REGION Network 38: Transition for STATE Num:43 Check Recovery
   RUNG wire#powerrail
      Contact( #s43_ChkRecovery )
      I_Contact( #sStWtResetRel )
      Contact( #sSst )
      wire#w1
      I_Contact( #iProcessOver )
      Coil( #s43_ChkRecovery_T1 )
   END_RUNG
   RUNG wire#w1
      I_Contact( #s43_ChkRecovery_T1 )
      Contact( #iProcessOver )
      Coil( #s43_ChkRecovery_T2 )
   END_RUNG
   // the same network as SCL:
   #_w1 := #s43_ChkRecovery AND NOT #sStWtResetRel AND #sSst;
   #s43_ChkRecovery_T1 := #_w1 AND NOT #iProcessOver;
   #s43_ChkRecovery_T2 := #_w1 AND NOT #s43_ChkRecovery_T1 AND #iProcessOver;
END_REGION

REGION Network 39: STATE Num:43 Check Recovery
   RUNG wire#powerrail
      Contact( #s43_ChkRecovery )
      wire#w1
      I_Contact( #sStWtResetRel )
      I_Contact( #s43_ChkRecovery_T1 )
      I_Contact( #s43_ChkRecovery_T2 )
      wire#w2
      Coil( #s43_ChkRecovery )
   END_RUNG
   RUNG wire#powerrail
      Contact( #s29_WaitProcStart_T1 )
   END_RUNG wire#w1
   RUNG wire#w2
      { S7_GenerateENO := "TRUE" } Move(in := 43, out1 => #StateNo)
   END_RUNG
   // the same network as SCL:
   #s43_ChkRecovery := (#s43_ChkRecovery OR #s29_WaitProcStart_T1) AND NOT #sStWtResetRel AND NOT #s43_ChkRecovery_T1 AND NOT #s43_ChkRecovery_T2;
   IF #s43_ChkRecovery THEN #StateNo := 43; END_IF;
END_REGION
END_FUNCTION_BLOCK

FUNCTION_BLOCK "PR_PC4005_Operator_DecisionV4_653444"   // FB2, LAD
VERSION : 0.1
// stored: AutoNumber true, IsIECCheckEnabled false, UDAEnableTagReadback false
   VAR_INPUT
      iAutoRunning : Bool;
      iOperatorAuthorizationPB : Bool;
      iPCAckZero : Bool;
      iPCBypass : Bool;
      iPCDataReadOver : Bool;
      iPCDataWriteOver : Bool;
      iPalletPresentAtStation : Bool;
      iProcessOver : Bool;
      iProcessStartFormPZR : Bool;
      iRejectPB : Bool;
      iResetMem : Bool;
      iReset_fault : Bool;
      iScanOver : Bool;
      iScanResultNok : Bool;
      iScanResultOk : Bool;
      iScannerBypass : Bool;
      iSstMode : Bool;
      iSstPB : Bool;
      iUnloadCycleSelection : Bool;
   END_VAR
   VAR_OUTPUT
      qPCReadCmd : Bool;
      qPCWriteCmd : Bool;
      qProcessOver : Bool;
      qResetPalletStatusData : Bool;
      qScanCmd : Bool;
   END_VAR
   VAR DB_SPECIFIC
      StateNo : Int;
      s29_WaitProcStart : Bool;
      s29_WaitProcStart_T1 : Bool;
      s30_WaitCartnSheetOp : Bool;
      s30_WaitCartnSheetOp_T1 : Bool;
      s31_ChkCycleSelect : Bool;
      s31_ChkCycleSelect_T1 : Bool;
      s31_ChkCycleSelect_T2 : Bool;
      s32_WaitScanOver : Bool;
      s32_WaitScanOver_T1 : Bool;
      s33_ChkScanResult : Bool;
      s33_ChkScanResult_T1 : Bool;
      s33_ChkScanResult_T2 : Bool;
      s34_WaitOpDecision : Bool;
      s34_WaitOpDecision_T1 : Bool;
      s34_WaitOpDecision_T2 : Bool;
      s35_ChkPCAckReset0 : Bool;
      s35_ChkPCAckReset0_T1 : Bool;
      s36_WaitDataReadPC : Bool;
      s36_WaitDataReadPC_T1 : Bool;
      s38_WaitProcStartLow : Bool;
      s38_WaitProcStartLow_T1 : Bool;
      s39_WaitPalletAbsnt : Bool;
      s39_WaitPalletAbsnt_T1 : Bool;
      s40_WaitFaultReset : Bool;
      s40_WaitFaultReset_T1 : Bool;
      s41_ChkPCAckReset0Up : Bool;
      s41_ChkPCAckReset0Up_T1 : Bool;
      s42_WaitDataUploadPC : Bool;
      s42_WaitDataUploadPC_T1 : Bool;
      s43_ChkRecovery : Bool;
      s43_ChkRecovery_T1 : Bool;
      s43_ChkRecovery_T2 : Bool;
      sPalletAccepted : Bool;
      sProcessOver : Bool;
      sSst : Bool;
      sSstPulse : Bool;
      sSstRise : Bool;
      sStWtResetRel : Bool;
      sStWtResetRel_T1 : Bool;
   END_VAR
   VAR_TEMP
      tOne : Bool;
   END_VAR
   VAR_TEMP   // added for the SCL form of the ladder/FBD networks
      _w1 : Bool;
   END_VAR
BEGIN

REGION Network 1
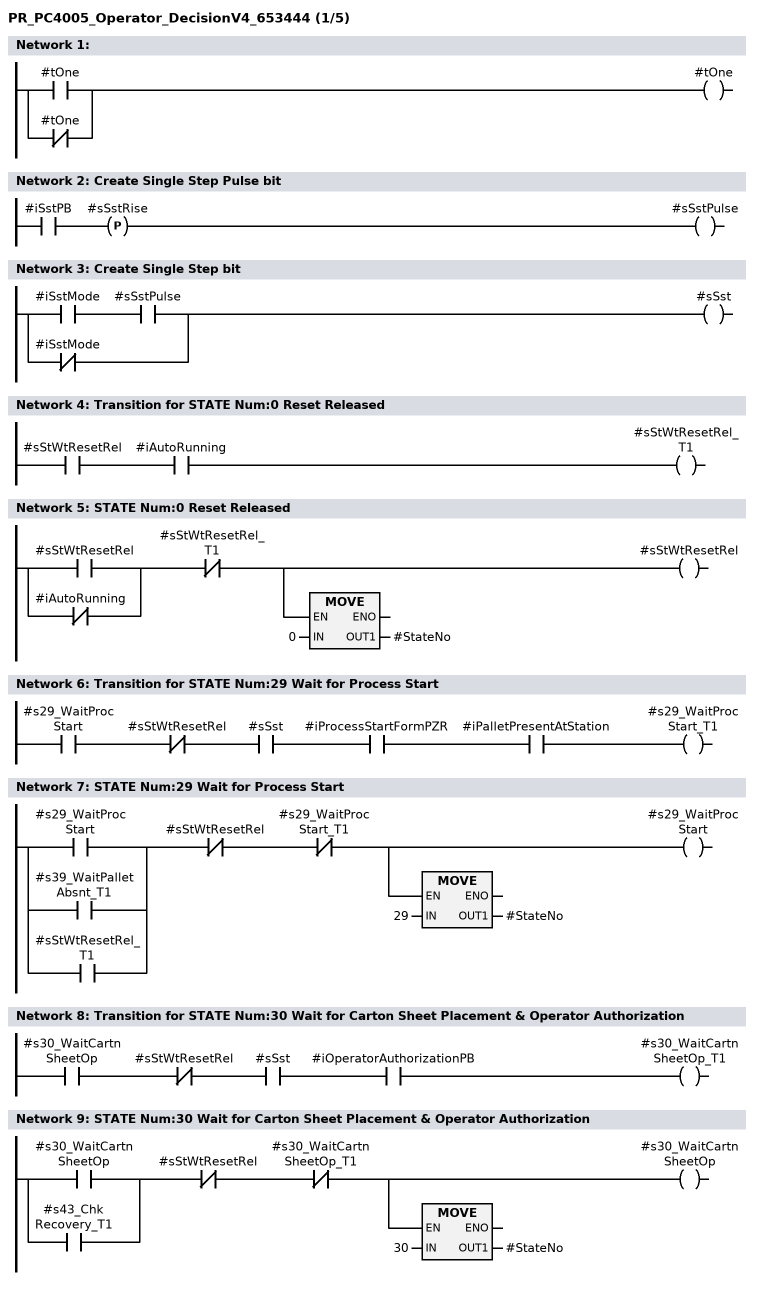
   RUNG wire#powerrail
      Contact( #tOne )
      wire#w1
      Coil( #tOne )
   END_RUNG
   RUNG wire#powerrail
      I_Contact( #tOne )
   END_RUNG wire#w1
   // the same network as SCL:
   #tOne := #tOne OR NOT #tOne;
END_REGION

REGION Network 2: Create Single Step Pulse bit
   RUNG wire#powerrail
      Contact( #iSstPB )
      P_Trig( #sSstRise )
      Coil( #sSstPulse )
   END_RUNG
   // the same network as SCL:
   #_w1 := #iSstPB AND NOT #sSstRise;   // rising edge
   #sSstRise := #iSstPB;
   #sSstPulse := #_w1;
END_REGION

REGION Network 3: Create Single Step bit
   RUNG wire#powerrail
      Contact( #iSstMode )
      Contact( #sSstPulse )
      wire#w1
      Coil( #sSst )
   END_RUNG
   RUNG wire#powerrail
      I_Contact( #iSstMode )
   END_RUNG wire#w1
   // the same network as SCL:
   #sSst := (#iSstMode AND #sSstPulse) OR NOT #iSstMode;
END_REGION

REGION Network 4: Transition for STATE Num:0 Reset Released
   RUNG wire#powerrail
      Contact( #sStWtResetRel )
      Contact( #iAutoRunning )
      Coil( #sStWtResetRel_T1 )
   END_RUNG
   // the same network as SCL:
   #sStWtResetRel_T1 := #sStWtResetRel AND #iAutoRunning;
END_REGION

REGION Network 5: STATE Num:0 Reset Released
   RUNG wire#powerrail
      Contact( #sStWtResetRel )
      wire#w1
      I_Contact( #sStWtResetRel_T1 )
      wire#w2
      Coil( #sStWtResetRel )
   END_RUNG
   RUNG wire#powerrail
      I_Contact( #iAutoRunning )
   END_RUNG wire#w1
   RUNG wire#w2
      { S7_GenerateENO := "TRUE" } Move(in := 0, out1 => #StateNo)
   END_RUNG
   // the same network as SCL:
   #sStWtResetRel := (#sStWtResetRel OR NOT #iAutoRunning) AND NOT #sStWtResetRel_T1;
   IF #sStWtResetRel THEN #StateNo := 0; END_IF;
END_REGION

REGION Network 6: Transition for STATE Num:29 Wait for Process Start
   RUNG wire#powerrail
      Contact( #s29_WaitProcStart )
      I_Contact( #sStWtResetRel )
      Contact( #sSst )
      Contact( #iProcessStartFormPZR )
      Contact( #iPalletPresentAtStation )
      Coil( #s29_WaitProcStart_T1 )
   END_RUNG
   // the same network as SCL:
   #s29_WaitProcStart_T1 := #s29_WaitProcStart AND NOT #sStWtResetRel AND #sSst AND #iProcessStartFormPZR AND #iPalletPresentAtStation;
END_REGION

REGION Network 7: STATE Num:29 Wait for Process Start
   RUNG wire#powerrail
      Contact( #s29_WaitProcStart )
      wire#w1
      I_Contact( #sStWtResetRel )
      I_Contact( #s29_WaitProcStart_T1 )
      wire#w2
      Coil( #s29_WaitProcStart )
   END_RUNG
   RUNG wire#powerrail
      Contact( #s39_WaitPalletAbsnt_T1 )
   END_RUNG wire#w1
   RUNG wire#powerrail
      Contact( #sStWtResetRel_T1 )
   END_RUNG wire#w1
   RUNG wire#w2
      { S7_GenerateENO := "TRUE" } Move(in := 29, out1 => #StateNo)
   END_RUNG
   // the same network as SCL:
   #s29_WaitProcStart := (#s29_WaitProcStart OR #s39_WaitPalletAbsnt_T1 OR #sStWtResetRel_T1) AND NOT #sStWtResetRel AND NOT #s29_WaitProcStart_T1;
   IF #s29_WaitProcStart THEN #StateNo := 29; END_IF;
END_REGION

REGION Network 8: Transition for STATE Num:30 Wait for Carton Sheet Placement & Operator Authorization
   RUNG wire#powerrail
      Contact( #s30_WaitCartnSheetOp )
      I_Contact( #sStWtResetRel )
      Contact( #sSst )
      Contact( #iOperatorAuthorizationPB )
      Coil( #s30_WaitCartnSheetOp_T1 )
   END_RUNG
   // the same network as SCL:
   #s30_WaitCartnSheetOp_T1 := #s30_WaitCartnSheetOp AND NOT #sStWtResetRel AND #sSst AND #iOperatorAuthorizationPB;
END_REGION

REGION Network 9: STATE Num:30 Wait for Carton Sheet Placement & Operator Authorization
   RUNG wire#powerrail
      Contact( #s30_WaitCartnSheetOp )
      wire#w1
      I_Contact( #sStWtResetRel )
      I_Contact( #s30_WaitCartnSheetOp_T1 )
      wire#w2
      Coil( #s30_WaitCartnSheetOp )
   END_RUNG
   RUNG wire#powerrail
      Contact( #s43_ChkRecovery_T1 )
   END_RUNG wire#w1
   RUNG wire#w2
      { S7_GenerateENO := "TRUE" } Move(in := 30, out1 => #StateNo)
   END_RUNG
   // the same network as SCL:
   #s30_WaitCartnSheetOp := (#s30_WaitCartnSheetOp OR #s43_ChkRecovery_T1) AND NOT #sStWtResetRel AND NOT #s30_WaitCartnSheetOp_T1;
   IF #s30_WaitCartnSheetOp THEN #StateNo := 30; END_IF;
END_REGION

REGION Network 10: Transition for STATE Num:31 Check Cycle Selection
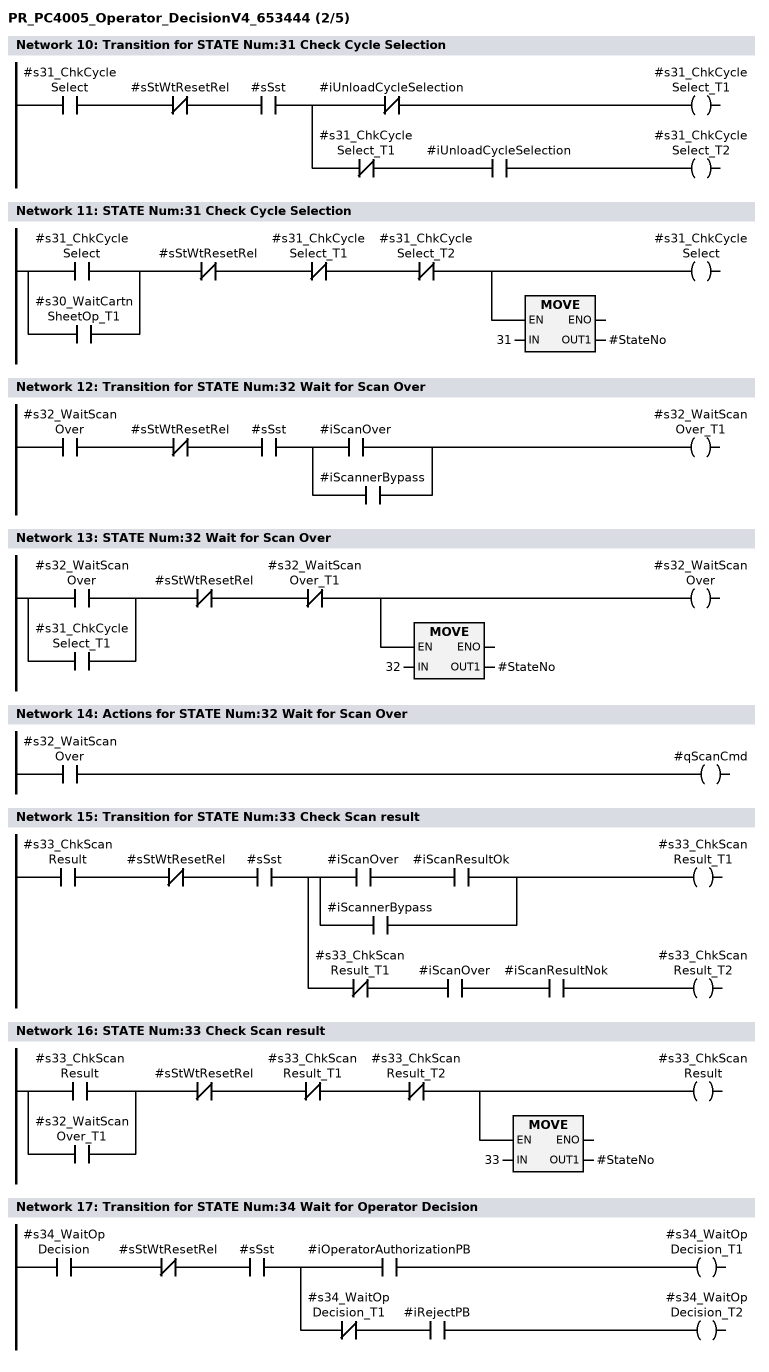
   RUNG wire#powerrail
      Contact( #s31_ChkCycleSelect )
      I_Contact( #sStWtResetRel )
      Contact( #sSst )
      wire#w1
      I_Contact( #iUnloadCycleSelection )
      Coil( #s31_ChkCycleSelect_T1 )
   END_RUNG
   RUNG wire#w1
      I_Contact( #s31_ChkCycleSelect_T1 )
      Contact( #iUnloadCycleSelection )
      Coil( #s31_ChkCycleSelect_T2 )
   END_RUNG
   // the same network as SCL:
   #_w1 := #s31_ChkCycleSelect AND NOT #sStWtResetRel AND #sSst;
   #s31_ChkCycleSelect_T1 := #_w1 AND NOT #iUnloadCycleSelection;
   #s31_ChkCycleSelect_T2 := #_w1 AND NOT #s31_ChkCycleSelect_T1 AND #iUnloadCycleSelection;
END_REGION

REGION Network 11: STATE Num:31 Check Cycle Selection
   RUNG wire#powerrail
      Contact( #s31_ChkCycleSelect )
      wire#w1
      I_Contact( #sStWtResetRel )
      I_Contact( #s31_ChkCycleSelect_T1 )
      I_Contact( #s31_ChkCycleSelect_T2 )
      wire#w2
      Coil( #s31_ChkCycleSelect )
   END_RUNG
   RUNG wire#powerrail
      Contact( #s30_WaitCartnSheetOp_T1 )
   END_RUNG wire#w1
   RUNG wire#w2
      { S7_GenerateENO := "TRUE" } Move(in := 31, out1 => #StateNo)
   END_RUNG
   // the same network as SCL:
   #s31_ChkCycleSelect := (#s31_ChkCycleSelect OR #s30_WaitCartnSheetOp_T1) AND NOT #sStWtResetRel AND NOT #s31_ChkCycleSelect_T1 AND NOT #s31_ChkCycleSelect_T2;
   IF #s31_ChkCycleSelect THEN #StateNo := 31; END_IF;
END_REGION

REGION Network 12: Transition for STATE Num:32 Wait for Scan Over
   RUNG wire#powerrail
      Contact( #s32_WaitScanOver )
      I_Contact( #sStWtResetRel )
      Contact( #sSst )
      wire#w1
      Contact( #iScanOver )
      wire#w2
      Coil( #s32_WaitScanOver_T1 )
   END_RUNG
   RUNG wire#w1
      Contact( #iScannerBypass )
   END_RUNG wire#w2
   // the same network as SCL:
   #s32_WaitScanOver_T1 := #s32_WaitScanOver AND NOT #sStWtResetRel AND #sSst AND (#iScanOver OR #iScannerBypass);
END_REGION

REGION Network 13: STATE Num:32 Wait for Scan Over
   RUNG wire#powerrail
      Contact( #s32_WaitScanOver )
      wire#w1
      I_Contact( #sStWtResetRel )
      I_Contact( #s32_WaitScanOver_T1 )
      wire#w2
      Coil( #s32_WaitScanOver )
   END_RUNG
   RUNG wire#powerrail
      Contact( #s31_ChkCycleSelect_T1 )
   END_RUNG wire#w1
   RUNG wire#w2
      { S7_GenerateENO := "TRUE" } Move(in := 32, out1 => #StateNo)
   END_RUNG
   // the same network as SCL:
   #s32_WaitScanOver := (#s32_WaitScanOver OR #s31_ChkCycleSelect_T1) AND NOT #sStWtResetRel AND NOT #s32_WaitScanOver_T1;
   IF #s32_WaitScanOver THEN #StateNo := 32; END_IF;
END_REGION

REGION Network 14: Actions for STATE Num:32 Wait for Scan Over
   RUNG wire#powerrail
      Contact( #s32_WaitScanOver )
      Coil( #qScanCmd )
   END_RUNG
   // the same network as SCL:
   #qScanCmd := #s32_WaitScanOver;
END_REGION

REGION Network 15: Transition for STATE Num:33 Check Scan result
   RUNG wire#powerrail
      Contact( #s33_ChkScanResult )
      I_Contact( #sStWtResetRel )
      Contact( #sSst )
      wire#w1
      Contact( #iScanOver )
      Contact( #iScanResultOk )
      wire#w2
      Coil( #s33_ChkScanResult_T1 )
   END_RUNG
   RUNG wire#w1
      Contact( #iScannerBypass )
   END_RUNG wire#w2
   RUNG wire#w1
      I_Contact( #s33_ChkScanResult_T1 )
      Contact( #iScanOver )
      Contact( #iScanResultNok )
      Coil( #s33_ChkScanResult_T2 )
   END_RUNG
   // the same network as SCL:
   #_w1 := #s33_ChkScanResult AND NOT #sStWtResetRel AND #sSst;
   #s33_ChkScanResult_T1 := #_w1 AND ((#iScanOver AND #iScanResultOk) OR #iScannerBypass);
   #s33_ChkScanResult_T2 := #_w1 AND NOT #s33_ChkScanResult_T1 AND #iScanOver AND #iScanResultNok;
END_REGION

REGION Network 16: STATE Num:33 Check Scan result
   RUNG wire#powerrail
      Contact( #s33_ChkScanResult )
      wire#w1
      I_Contact( #sStWtResetRel )
      I_Contact( #s33_ChkScanResult_T1 )
      I_Contact( #s33_ChkScanResult_T2 )
      wire#w2
      Coil( #s33_ChkScanResult )
   END_RUNG
   RUNG wire#powerrail
      Contact( #s32_WaitScanOver_T1 )
   END_RUNG wire#w1
   RUNG wire#w2
      { S7_GenerateENO := "TRUE" } Move(in := 33, out1 => #StateNo)
   END_RUNG
   // the same network as SCL:
   #s33_ChkScanResult := (#s33_ChkScanResult OR #s32_WaitScanOver_T1) AND NOT #sStWtResetRel AND NOT #s33_ChkScanResult_T1 AND NOT #s33_ChkScanResult_T2;
   IF #s33_ChkScanResult THEN #StateNo := 33; END_IF;
END_REGION

REGION Network 17: Transition for STATE Num:34 Wait for Operator Decision
   RUNG wire#powerrail
      Contact( #s34_WaitOpDecision )
      I_Contact( #sStWtResetRel )
      Contact( #sSst )
      wire#w1
      Contact( #iOperatorAuthorizationPB )
      Coil( #s34_WaitOpDecision_T1 )
   END_RUNG
   RUNG wire#w1
      I_Contact( #s34_WaitOpDecision_T1 )
      Contact( #iRejectPB )
      Coil( #s34_WaitOpDecision_T2 )
   END_RUNG
   // the same network as SCL:
   #_w1 := #s34_WaitOpDecision AND NOT #sStWtResetRel AND #sSst;
   #s34_WaitOpDecision_T1 := #_w1 AND #iOperatorAuthorizationPB;
   #s34_WaitOpDecision_T2 := #_w1 AND NOT #s34_WaitOpDecision_T1 AND #iRejectPB;
END_REGION

REGION Network 18: STATE Num:34 Wait for Operator Decision
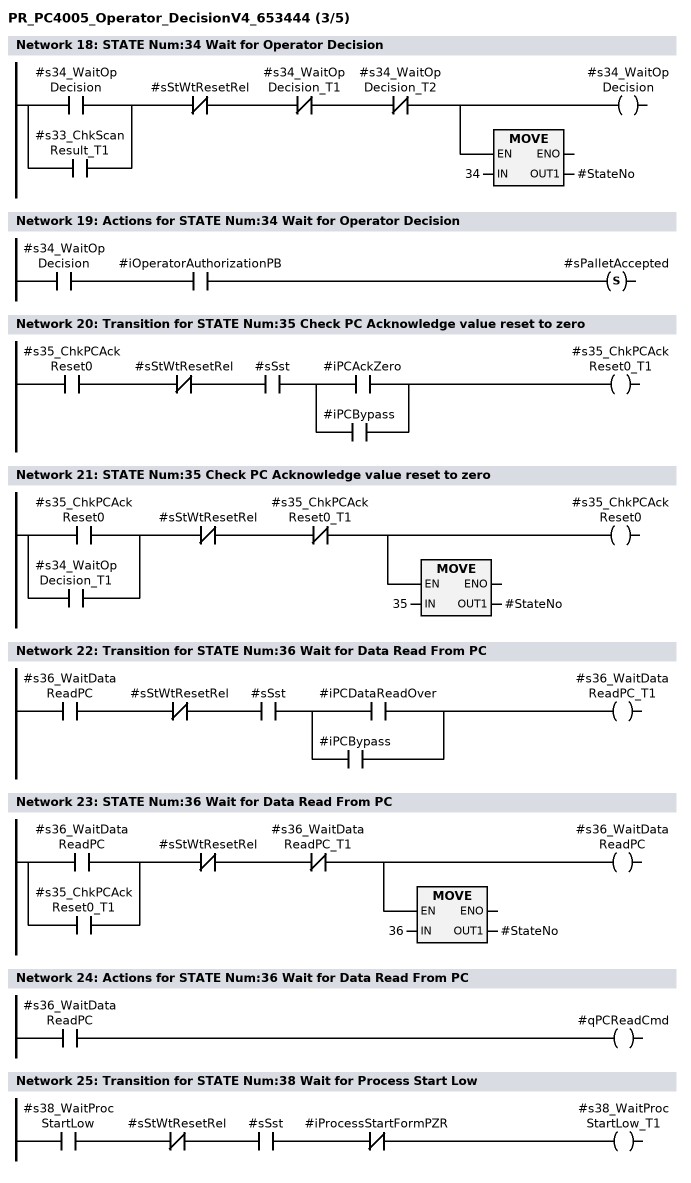
   RUNG wire#powerrail
      Contact( #s34_WaitOpDecision )
      wire#w1
      I_Contact( #sStWtResetRel )
      I_Contact( #s34_WaitOpDecision_T1 )
      I_Contact( #s34_WaitOpDecision_T2 )
      wire#w2
      Coil( #s34_WaitOpDecision )
   END_RUNG
   RUNG wire#powerrail
      Contact( #s33_ChkScanResult_T1 )
   END_RUNG wire#w1
   RUNG wire#w2
      { S7_GenerateENO := "TRUE" } Move(in := 34, out1 => #StateNo)
   END_RUNG
   // the same network as SCL:
   #s34_WaitOpDecision := (#s34_WaitOpDecision OR #s33_ChkScanResult_T1) AND NOT #sStWtResetRel AND NOT #s34_WaitOpDecision_T1 AND NOT #s34_WaitOpDecision_T2;
   IF #s34_WaitOpDecision THEN #StateNo := 34; END_IF;
END_REGION

REGION Network 19: Actions for STATE Num:34 Wait for Operator Decision
   RUNG wire#powerrail
      Contact( #s34_WaitOpDecision )
      Contact( #iOperatorAuthorizationPB )
      S_Coil( #sPalletAccepted )
   END_RUNG
   // the same network as SCL:
   IF #s34_WaitOpDecision AND #iOperatorAuthorizationPB THEN #sPalletAccepted := TRUE; END_IF;
END_REGION

REGION Network 20: Transition for STATE Num:35 Check PC Acknowledge value reset to zero
   RUNG wire#powerrail
      Contact( #s35_ChkPCAckReset0 )
      I_Contact( #sStWtResetRel )
      Contact( #sSst )
      wire#w1
      Contact( #iPCAckZero )
      wire#w2
      Coil( #s35_ChkPCAckReset0_T1 )
   END_RUNG
   RUNG wire#w1
      Contact( #iPCBypass )
   END_RUNG wire#w2
   // the same network as SCL:
   #s35_ChkPCAckReset0_T1 := #s35_ChkPCAckReset0 AND NOT #sStWtResetRel AND #sSst AND (#iPCAckZero OR #iPCBypass);
END_REGION

REGION Network 21: STATE Num:35 Check PC Acknowledge value reset to zero
   RUNG wire#powerrail
      Contact( #s35_ChkPCAckReset0 )
      wire#w1
      I_Contact( #sStWtResetRel )
      I_Contact( #s35_ChkPCAckReset0_T1 )
      wire#w2
      Coil( #s35_ChkPCAckReset0 )
   END_RUNG
   RUNG wire#powerrail
      Contact( #s34_WaitOpDecision_T1 )
   END_RUNG wire#w1
   RUNG wire#w2
      { S7_GenerateENO := "TRUE" } Move(in := 35, out1 => #StateNo)
   END_RUNG
   // the same network as SCL:
   #s35_ChkPCAckReset0 := (#s35_ChkPCAckReset0 OR #s34_WaitOpDecision_T1) AND NOT #sStWtResetRel AND NOT #s35_ChkPCAckReset0_T1;
   IF #s35_ChkPCAckReset0 THEN #StateNo := 35; END_IF;
END_REGION

REGION Network 22: Transition for STATE Num:36 Wait for Data Read From PC
   RUNG wire#powerrail
      Contact( #s36_WaitDataReadPC )
      I_Contact( #sStWtResetRel )
      Contact( #sSst )
      wire#w1
      Contact( #iPCDataReadOver )
      wire#w2
      Coil( #s36_WaitDataReadPC_T1 )
   END_RUNG
   RUNG wire#w1
      Contact( #iPCBypass )
   END_RUNG wire#w2
   // the same network as SCL:
   #s36_WaitDataReadPC_T1 := #s36_WaitDataReadPC AND NOT #sStWtResetRel AND #sSst AND (#iPCDataReadOver OR #iPCBypass);
END_REGION

REGION Network 23: STATE Num:36 Wait for Data Read From PC
   RUNG wire#powerrail
      Contact( #s36_WaitDataReadPC )
      wire#w1
      I_Contact( #sStWtResetRel )
      I_Contact( #s36_WaitDataReadPC_T1 )
      wire#w2
      Coil( #s36_WaitDataReadPC )
   END_RUNG
   RUNG wire#powerrail
      Contact( #s35_ChkPCAckReset0_T1 )
   END_RUNG wire#w1
   RUNG wire#w2
      { S7_GenerateENO := "TRUE" } Move(in := 36, out1 => #StateNo)
   END_RUNG
   // the same network as SCL:
   #s36_WaitDataReadPC := (#s36_WaitDataReadPC OR #s35_ChkPCAckReset0_T1) AND NOT #sStWtResetRel AND NOT #s36_WaitDataReadPC_T1;
   IF #s36_WaitDataReadPC THEN #StateNo := 36; END_IF;
END_REGION

REGION Network 24: Actions for STATE Num:36 Wait for Data Read From PC
   RUNG wire#powerrail
      Contact( #s36_WaitDataReadPC )
      Coil( #qPCReadCmd )
   END_RUNG
   // the same network as SCL:
   #qPCReadCmd := #s36_WaitDataReadPC;
END_REGION

REGION Network 25: Transition for STATE Num:38 Wait for Process Start Low
   RUNG wire#powerrail
      Contact( #s38_WaitProcStartLow )
      I_Contact( #sStWtResetRel )
      Contact( #sSst )
      I_Contact( #iProcessStartFormPZR )
      Coil( #s38_WaitProcStartLow_T1 )
   END_RUNG
   // the same network as SCL:
   #s38_WaitProcStartLow_T1 := #s38_WaitProcStartLow AND NOT #sStWtResetRel AND #sSst AND NOT #iProcessStartFormPZR;
END_REGION

REGION Network 26: STATE Num:38 Wait for Process Start Low
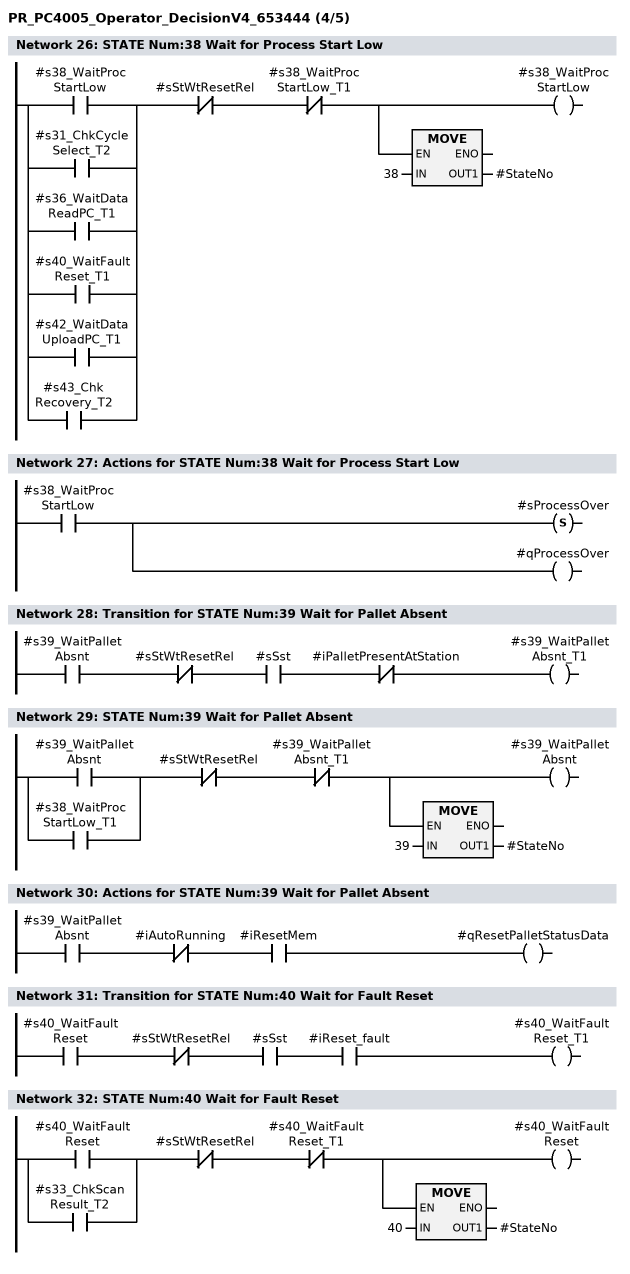
   RUNG wire#powerrail
      Contact( #s38_WaitProcStartLow )
      wire#w1
      I_Contact( #sStWtResetRel )
      I_Contact( #s38_WaitProcStartLow_T1 )
      wire#w2
      Coil( #s38_WaitProcStartLow )
   END_RUNG
   RUNG wire#powerrail
      Contact( #s31_ChkCycleSelect_T2 )
   END_RUNG wire#w1
   RUNG wire#powerrail
      Contact( #s36_WaitDataReadPC_T1 )
   END_RUNG wire#w1
   RUNG wire#powerrail
      Contact( #s40_WaitFaultReset_T1 )
   END_RUNG wire#w1
   RUNG wire#powerrail
      Contact( #s42_WaitDataUploadPC_T1 )
   END_RUNG wire#w1
   RUNG wire#powerrail
      Contact( #s43_ChkRecovery_T2 )
   END_RUNG wire#w1
   RUNG wire#w2
      { S7_GenerateENO := "TRUE" } Move(in := 38, out1 => #StateNo)
   END_RUNG
   // the same network as SCL:
   #s38_WaitProcStartLow := (#s38_WaitProcStartLow OR #s31_ChkCycleSelect_T2 OR #s36_WaitDataReadPC_T1 OR #s40_WaitFaultReset_T1 OR #s42_WaitDataUploadPC_T1 OR #s43_ChkRecovery_T2) AND NOT #sStWtResetRel AND NOT #s38_WaitProcStartLow_T1;
   IF #s38_WaitProcStartLow THEN #StateNo := 38; END_IF;
END_REGION

REGION Network 27: Actions for STATE Num:38 Wait for Process Start Low
   RUNG wire#powerrail
      Contact( #s38_WaitProcStartLow )
      wire#w1
      S_Coil( #sProcessOver )
   END_RUNG
   RUNG wire#w1
      Coil( #qProcessOver )
   END_RUNG
   // the same network as SCL:
   IF #s38_WaitProcStartLow THEN #sProcessOver := TRUE; END_IF;
   #qProcessOver := #s38_WaitProcStartLow;
END_REGION

REGION Network 28: Transition for STATE Num:39 Wait for Pallet Absent
   RUNG wire#powerrail
      Contact( #s39_WaitPalletAbsnt )
      I_Contact( #sStWtResetRel )
      Contact( #sSst )
      I_Contact( #iPalletPresentAtStation )
      Coil( #s39_WaitPalletAbsnt_T1 )
   END_RUNG
   // the same network as SCL:
   #s39_WaitPalletAbsnt_T1 := #s39_WaitPalletAbsnt AND NOT #sStWtResetRel AND #sSst AND NOT #iPalletPresentAtStation;
END_REGION

REGION Network 29: STATE Num:39 Wait for Pallet Absent
   RUNG wire#powerrail
      Contact( #s39_WaitPalletAbsnt )
      wire#w1
      I_Contact( #sStWtResetRel )
      I_Contact( #s39_WaitPalletAbsnt_T1 )
      wire#w2
      Coil( #s39_WaitPalletAbsnt )
   END_RUNG
   RUNG wire#powerrail
      Contact( #s38_WaitProcStartLow_T1 )
   END_RUNG wire#w1
   RUNG wire#w2
      { S7_GenerateENO := "TRUE" } Move(in := 39, out1 => #StateNo)
   END_RUNG
   // the same network as SCL:
   #s39_WaitPalletAbsnt := (#s39_WaitPalletAbsnt OR #s38_WaitProcStartLow_T1) AND NOT #sStWtResetRel AND NOT #s39_WaitPalletAbsnt_T1;
   IF #s39_WaitPalletAbsnt THEN #StateNo := 39; END_IF;
END_REGION

REGION Network 30: Actions for STATE Num:39 Wait for Pallet Absent
   RUNG wire#powerrail
      Contact( #s39_WaitPalletAbsnt )
      I_Contact( #iAutoRunning )
      Contact( #iResetMem )
      Coil( #qResetPalletStatusData )
   END_RUNG
   // the same network as SCL:
   #qResetPalletStatusData := #s39_WaitPalletAbsnt AND NOT #iAutoRunning AND #iResetMem;
END_REGION

REGION Network 31: Transition for STATE Num:40 Wait for Fault Reset
   RUNG wire#powerrail
      Contact( #s40_WaitFaultReset )
      I_Contact( #sStWtResetRel )
      Contact( #sSst )
      Contact( #iReset_fault )
      Coil( #s40_WaitFaultReset_T1 )
   END_RUNG
   // the same network as SCL:
   #s40_WaitFaultReset_T1 := #s40_WaitFaultReset AND NOT #sStWtResetRel AND #sSst AND #iReset_fault;
END_REGION

REGION Network 32: STATE Num:40 Wait for Fault Reset
   RUNG wire#powerrail
      Contact( #s40_WaitFaultReset )
      wire#w1
      I_Contact( #sStWtResetRel )
      I_Contact( #s40_WaitFaultReset_T1 )
      wire#w2
      Coil( #s40_WaitFaultReset )
   END_RUNG
   RUNG wire#powerrail
      Contact( #s33_ChkScanResult_T2 )
   END_RUNG wire#w1
   RUNG wire#w2
      { S7_GenerateENO := "TRUE" } Move(in := 40, out1 => #StateNo)
   END_RUNG
   // the same network as SCL:
   #s40_WaitFaultReset := (#s40_WaitFaultReset OR #s33_ChkScanResult_T2) AND NOT #sStWtResetRel AND NOT #s40_WaitFaultReset_T1;
   IF #s40_WaitFaultReset THEN #StateNo := 40; END_IF;
END_REGION

REGION Network 33: Transition for STATE Num:41 Check PC Acknowledge value reset to zero for Upload
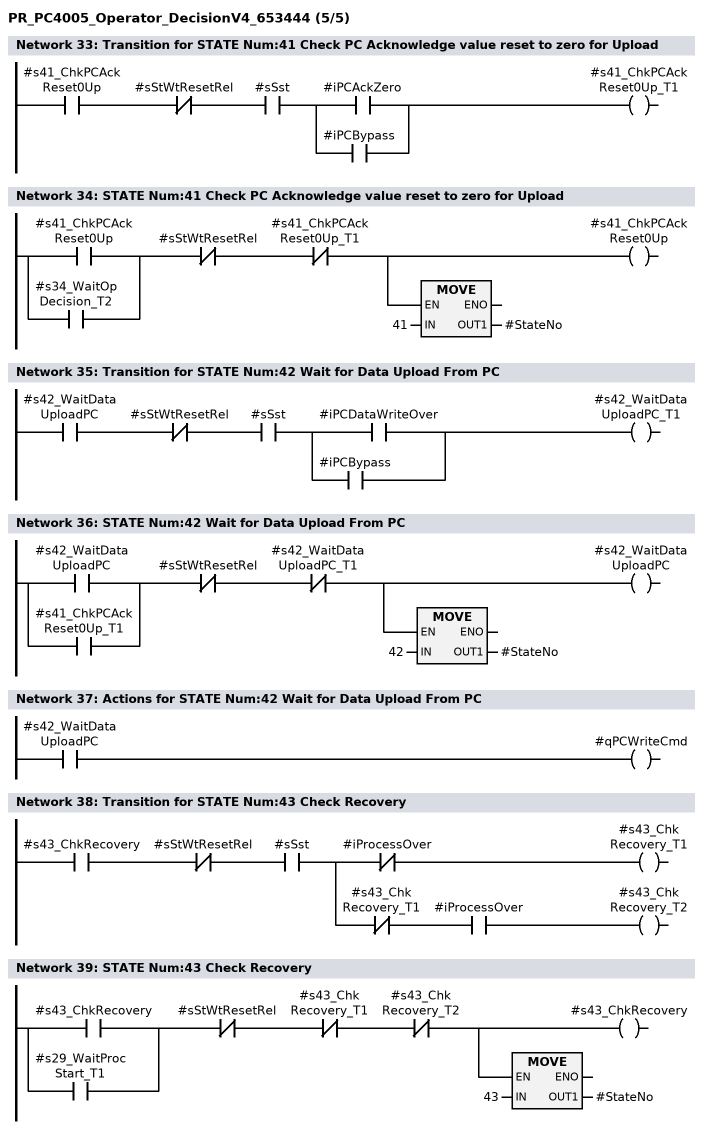
   RUNG wire#powerrail
      Contact( #s41_ChkPCAckReset0Up )
      I_Contact( #sStWtResetRel )
      Contact( #sSst )
      wire#w1
      Contact( #iPCAckZero )
      wire#w2
      Coil( #s41_ChkPCAckReset0Up_T1 )
   END_RUNG
   RUNG wire#w1
      Contact( #iPCBypass )
   END_RUNG wire#w2
   // the same network as SCL:
   #s41_ChkPCAckReset0Up_T1 := #s41_ChkPCAckReset0Up AND NOT #sStWtResetRel AND #sSst AND (#iPCAckZero OR #iPCBypass);
END_REGION

REGION Network 34: STATE Num:41 Check PC Acknowledge value reset to zero for Upload
   RUNG wire#powerrail
      Contact( #s41_ChkPCAckReset0Up )
      wire#w1
      I_Contact( #sStWtResetRel )
      I_Contact( #s41_ChkPCAckReset0Up_T1 )
      wire#w2
      Coil( #s41_ChkPCAckReset0Up )
   END_RUNG
   RUNG wire#powerrail
      Contact( #s34_WaitOpDecision_T2 )
   END_RUNG wire#w1
   RUNG wire#w2
      { S7_GenerateENO := "TRUE" } Move(in := 41, out1 => #StateNo)
   END_RUNG
   // the same network as SCL:
   #s41_ChkPCAckReset0Up := (#s41_ChkPCAckReset0Up OR #s34_WaitOpDecision_T2) AND NOT #sStWtResetRel AND NOT #s41_ChkPCAckReset0Up_T1;
   IF #s41_ChkPCAckReset0Up THEN #StateNo := 41; END_IF;
END_REGION

REGION Network 35: Transition for STATE Num:42 Wait for Data Upload From PC
   RUNG wire#powerrail
      Contact( #s42_WaitDataUploadPC )
      I_Contact( #sStWtResetRel )
      Contact( #sSst )
      wire#w1
      Contact( #iPCDataWriteOver )
      wire#w2
      Coil( #s42_WaitDataUploadPC_T1 )
   END_RUNG
   RUNG wire#w1
      Contact( #iPCBypass )
   END_RUNG wire#w2
   // the same network as SCL:
   #s42_WaitDataUploadPC_T1 := #s42_WaitDataUploadPC AND NOT #sStWtResetRel AND #sSst AND (#iPCDataWriteOver OR #iPCBypass);
END_REGION

REGION Network 36: STATE Num:42 Wait for Data Upload From PC
   RUNG wire#powerrail
      Contact( #s42_WaitDataUploadPC )
      wire#w1
      I_Contact( #sStWtResetRel )
      I_Contact( #s42_WaitDataUploadPC_T1 )
      wire#w2
      Coil( #s42_WaitDataUploadPC )
   END_RUNG
   RUNG wire#powerrail
      Contact( #s41_ChkPCAckReset0Up_T1 )
   END_RUNG wire#w1
   RUNG wire#w2
      { S7_GenerateENO := "TRUE" } Move(in := 42, out1 => #StateNo)
   END_RUNG
   // the same network as SCL:
   #s42_WaitDataUploadPC := (#s42_WaitDataUploadPC OR #s41_ChkPCAckReset0Up_T1) AND NOT #sStWtResetRel AND NOT #s42_WaitDataUploadPC_T1;
   IF #s42_WaitDataUploadPC THEN #StateNo := 42; END_IF;
END_REGION

REGION Network 37: Actions for STATE Num:42 Wait for Data Upload From PC
   RUNG wire#powerrail
      Contact( #s42_WaitDataUploadPC )
      Coil( #qPCWriteCmd )
   END_RUNG
   // the same network as SCL:
   #qPCWriteCmd := #s42_WaitDataUploadPC;
END_REGION

REGION Network 38: Transition for STATE Num:43 Check Recovery
   RUNG wire#powerrail
      Contact( #s43_ChkRecovery )
      I_Contact( #sStWtResetRel )
      Contact( #sSst )
      wire#w1
      I_Contact( #iProcessOver )
      Coil( #s43_ChkRecovery_T1 )
   END_RUNG
   RUNG wire#w1
      I_Contact( #s43_ChkRecovery_T1 )
      Contact( #iProcessOver )
      Coil( #s43_ChkRecovery_T2 )
   END_RUNG
   // the same network as SCL:
   #_w1 := #s43_ChkRecovery AND NOT #sStWtResetRel AND #sSst;
   #s43_ChkRecovery_T1 := #_w1 AND NOT #iProcessOver;
   #s43_ChkRecovery_T2 := #_w1 AND NOT #s43_ChkRecovery_T1 AND #iProcessOver;
END_REGION

REGION Network 39: STATE Num:43 Check Recovery
   RUNG wire#powerrail
      Contact( #s43_ChkRecovery )
      wire#w1
      I_Contact( #sStWtResetRel )
      I_Contact( #s43_ChkRecovery_T1 )
      I_Contact( #s43_ChkRecovery_T2 )
      wire#w2
      Coil( #s43_ChkRecovery )
   END_RUNG
   RUNG wire#powerrail
      Contact( #s29_WaitProcStart_T1 )
   END_RUNG wire#w1
   RUNG wire#w2
      { S7_GenerateENO := "TRUE" } Move(in := 43, out1 => #StateNo)
   END_RUNG
   // the same network as SCL:
   #s43_ChkRecovery := (#s43_ChkRecovery OR #s29_WaitProcStart_T1) AND NOT #sStWtResetRel AND NOT #s43_ChkRecovery_T1 AND NOT #s43_ChkRecovery_T2;
   IF #s43_ChkRecovery THEN #StateNo := 43; END_IF;
END_REGION
END_FUNCTION_BLOCK

FUNCTION_BLOCK "PR_PC4005_Operator_DecisionV4_77a371"   // FB1, LAD
VERSION : 0.1
// stored: AutoNumber true, IsIECCheckEnabled false, UDAEnableTagReadback false
   VAR_INPUT
      iAutoRunning : Bool;
      iOperatorAuthorizationPB : Bool;
      iPCAckZero : Bool;
      iPCBypass : Bool;
      iPCDataReadOver : Bool;
      iPCDataWriteOver : Bool;
      iPalletPresentAtStation : Bool;
      iProcessOver : Bool;
      iProcessStartFormPZR : Bool;
      iRejectPB : Bool;
      iResetMem : Bool;
      iReset_fault : Bool;
      iScanOver : Bool;
      iScanResultNok : Bool;
      iScanResultOk : Bool;
      iScannerBypass : Bool;
      iSstMode : Bool;
      iSstPB : Bool;
      iUnloadCycleSelection : Bool;
   END_VAR
   VAR_OUTPUT
      qPCReadCmd : Bool;
      qPCWriteCmd : Bool;
      qProcessOver : Bool;
      qResetPalletStatusData : Bool;
      qScanCmd : Bool;
   END_VAR
   VAR DB_SPECIFIC
      StateNo : Int;
      s29_WaitProcStart : Bool;
      s29_WaitProcStart_T1 : Bool;
      s30_WaitCartnSheetOp : Bool;
      s30_WaitCartnSheetOp_T1 : Bool;
      s31_ChkCycleSelect : Bool;
      s31_ChkCycleSelect_T1 : Bool;
      s31_ChkCycleSelect_T2 : Bool;
      s32_WaitScanOver : Bool;
      s32_WaitScanOver_T1 : Bool;
      s33_ChkScanResult : Bool;
      s33_ChkScanResult_T1 : Bool;
      s33_ChkScanResult_T2 : Bool;
      s34_WaitOpDecision : Bool;
      s34_WaitOpDecision_T1 : Bool;
      s34_WaitOpDecision_T2 : Bool;
      s35_ChkPCAckReset0 : Bool;
      s35_ChkPCAckReset0_T1 : Bool;
      s36_WaitDataReadPC : Bool;
      s36_WaitDataReadPC_T1 : Bool;
      s38_WaitProcStartLow : Bool;
      s38_WaitProcStartLow_T1 : Bool;
      s39_WaitPalletAbsnt : Bool;
      s39_WaitPalletAbsnt_T1 : Bool;
      s40_WaitFaultReset : Bool;
      s40_WaitFaultReset_T1 : Bool;
      s41_ChkPCAckReset0Up : Bool;
      s41_ChkPCAckReset0Up_T1 : Bool;
      s42_WaitDataUploadPC : Bool;
      s42_WaitDataUploadPC_T1 : Bool;
      s43_ChkRecovery : Bool;
      s43_ChkRecovery_T1 : Bool;
      s43_ChkRecovery_T2 : Bool;
      sPalletAccepted : Bool;
      sProcessOver : Bool;
      sSst : Bool;
      sSstPulse : Bool;
      sSstRise : Bool;
      sStWtResetRel : Bool;
      sStWtResetRel_T1 : Bool;
   END_VAR
   VAR_TEMP
      tOne : Bool;
   END_VAR
   VAR_TEMP   // added for the SCL form of the ladder/FBD networks
      _w1 : Bool;
   END_VAR
BEGIN

REGION Network 1
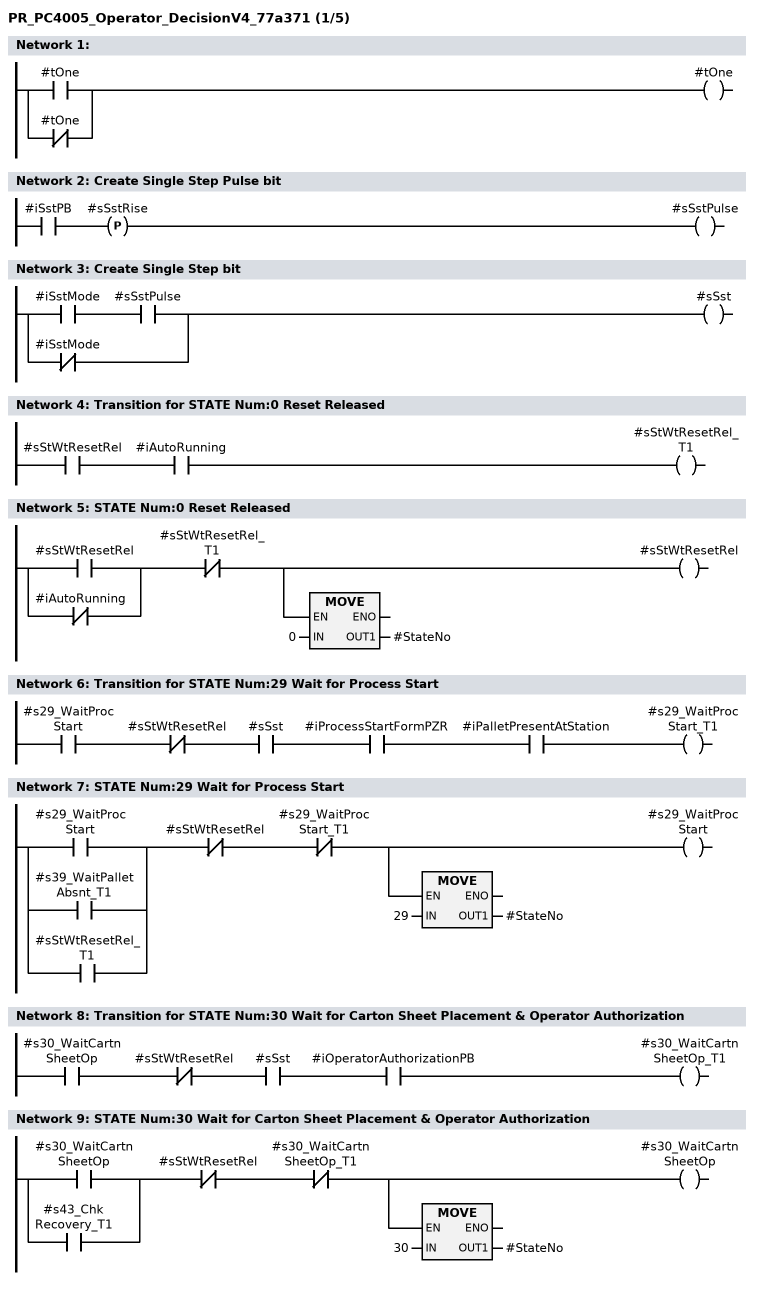
   RUNG wire#powerrail
      Contact( #tOne )
      wire#w1
      Coil( #tOne )
   END_RUNG
   RUNG wire#powerrail
      I_Contact( #tOne )
   END_RUNG wire#w1
   // the same network as SCL:
   #tOne := #tOne OR NOT #tOne;
END_REGION

REGION Network 2: Create Single Step Pulse bit
   RUNG wire#powerrail
      Contact( #iSstPB )
      P_Trig( #sSstRise )
      Coil( #sSstPulse )
   END_RUNG
   // the same network as SCL:
   #_w1 := #iSstPB AND NOT #sSstRise;   // rising edge
   #sSstRise := #iSstPB;
   #sSstPulse := #_w1;
END_REGION

REGION Network 3: Create Single Step bit
   RUNG wire#powerrail
      Contact( #iSstMode )
      Contact( #sSstPulse )
      wire#w1
      Coil( #sSst )
   END_RUNG
   RUNG wire#powerrail
      I_Contact( #iSstMode )
   END_RUNG wire#w1
   // the same network as SCL:
   #sSst := (#iSstMode AND #sSstPulse) OR NOT #iSstMode;
END_REGION

REGION Network 4: Transition for STATE Num:0 Reset Released
   RUNG wire#powerrail
      Contact( #sStWtResetRel )
      Contact( #iAutoRunning )
      Coil( #sStWtResetRel_T1 )
   END_RUNG
   // the same network as SCL:
   #sStWtResetRel_T1 := #sStWtResetRel AND #iAutoRunning;
END_REGION

REGION Network 5: STATE Num:0 Reset Released
   RUNG wire#powerrail
      Contact( #sStWtResetRel )
      wire#w1
      I_Contact( #sStWtResetRel_T1 )
      wire#w2
      Coil( #sStWtResetRel )
   END_RUNG
   RUNG wire#powerrail
      I_Contact( #iAutoRunning )
   END_RUNG wire#w1
   RUNG wire#w2
      { S7_GenerateENO := "TRUE" } Move(in := 0, out1 => #StateNo)
   END_RUNG
   // the same network as SCL:
   #sStWtResetRel := (#sStWtResetRel OR NOT #iAutoRunning) AND NOT #sStWtResetRel_T1;
   IF #sStWtResetRel THEN #StateNo := 0; END_IF;
END_REGION

REGION Network 6: Transition for STATE Num:29 Wait for Process Start
   RUNG wire#powerrail
      Contact( #s29_WaitProcStart )
      I_Contact( #sStWtResetRel )
      Contact( #sSst )
      Contact( #iProcessStartFormPZR )
      Contact( #iPalletPresentAtStation )
      Coil( #s29_WaitProcStart_T1 )
   END_RUNG
   // the same network as SCL:
   #s29_WaitProcStart_T1 := #s29_WaitProcStart AND NOT #sStWtResetRel AND #sSst AND #iProcessStartFormPZR AND #iPalletPresentAtStation;
END_REGION

REGION Network 7: STATE Num:29 Wait for Process Start
   RUNG wire#powerrail
      Contact( #s29_WaitProcStart )
      wire#w1
      I_Contact( #sStWtResetRel )
      I_Contact( #s29_WaitProcStart_T1 )
      wire#w2
      Coil( #s29_WaitProcStart )
   END_RUNG
   RUNG wire#powerrail
      Contact( #s39_WaitPalletAbsnt_T1 )
   END_RUNG wire#w1
   RUNG wire#powerrail
      Contact( #sStWtResetRel_T1 )
   END_RUNG wire#w1
   RUNG wire#w2
      { S7_GenerateENO := "TRUE" } Move(in := 29, out1 => #StateNo)
   END_RUNG
   // the same network as SCL:
   #s29_WaitProcStart := (#s29_WaitProcStart OR #s39_WaitPalletAbsnt_T1 OR #sStWtResetRel_T1) AND NOT #sStWtResetRel AND NOT #s29_WaitProcStart_T1;
   IF #s29_WaitProcStart THEN #StateNo := 29; END_IF;
END_REGION

REGION Network 8: Transition for STATE Num:30 Wait for Carton Sheet Placement & Operator Authorization
   RUNG wire#powerrail
      Contact( #s30_WaitCartnSheetOp )
      I_Contact( #sStWtResetRel )
      Contact( #sSst )
      Contact( #iOperatorAuthorizationPB )
      Coil( #s30_WaitCartnSheetOp_T1 )
   END_RUNG
   // the same network as SCL:
   #s30_WaitCartnSheetOp_T1 := #s30_WaitCartnSheetOp AND NOT #sStWtResetRel AND #sSst AND #iOperatorAuthorizationPB;
END_REGION

REGION Network 9: STATE Num:30 Wait for Carton Sheet Placement & Operator Authorization
   RUNG wire#powerrail
      Contact( #s30_WaitCartnSheetOp )
      wire#w1
      I_Contact( #sStWtResetRel )
      I_Contact( #s30_WaitCartnSheetOp_T1 )
      wire#w2
      Coil( #s30_WaitCartnSheetOp )
   END_RUNG
   RUNG wire#powerrail
      Contact( #s43_ChkRecovery_T1 )
   END_RUNG wire#w1
   RUNG wire#w2
      { S7_GenerateENO := "TRUE" } Move(in := 30, out1 => #StateNo)
   END_RUNG
   // the same network as SCL:
   #s30_WaitCartnSheetOp := (#s30_WaitCartnSheetOp OR #s43_ChkRecovery_T1) AND NOT #sStWtResetRel AND NOT #s30_WaitCartnSheetOp_T1;
   IF #s30_WaitCartnSheetOp THEN #StateNo := 30; END_IF;
END_REGION

REGION Network 10: Transition for STATE Num:31 Check Cycle Selection
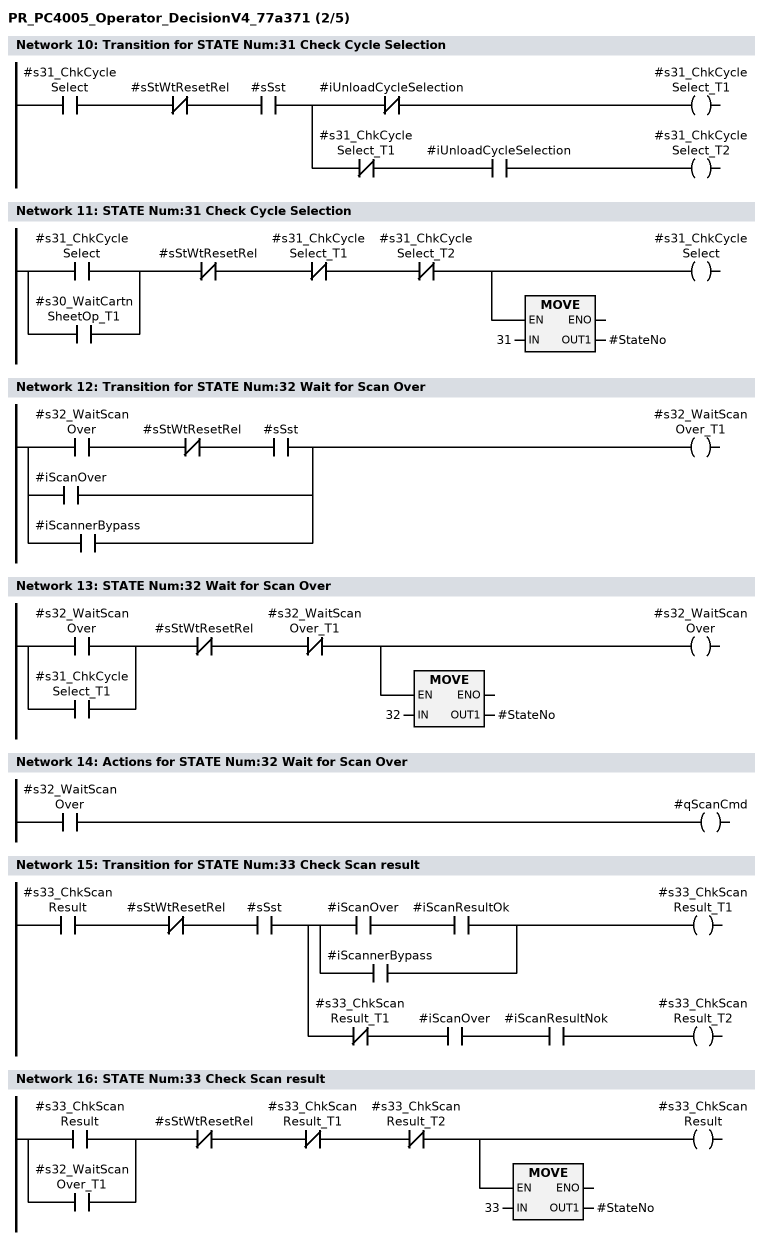
   RUNG wire#powerrail
      Contact( #s31_ChkCycleSelect )
      I_Contact( #sStWtResetRel )
      Contact( #sSst )
      wire#w1
      I_Contact( #iUnloadCycleSelection )
      Coil( #s31_ChkCycleSelect_T1 )
   END_RUNG
   RUNG wire#w1
      I_Contact( #s31_ChkCycleSelect_T1 )
      Contact( #iUnloadCycleSelection )
      Coil( #s31_ChkCycleSelect_T2 )
   END_RUNG
   // the same network as SCL:
   #_w1 := #s31_ChkCycleSelect AND NOT #sStWtResetRel AND #sSst;
   #s31_ChkCycleSelect_T1 := #_w1 AND NOT #iUnloadCycleSelection;
   #s31_ChkCycleSelect_T2 := #_w1 AND NOT #s31_ChkCycleSelect_T1 AND #iUnloadCycleSelection;
END_REGION

REGION Network 11: STATE Num:31 Check Cycle Selection
   RUNG wire#powerrail
      Contact( #s31_ChkCycleSelect )
      wire#w1
      I_Contact( #sStWtResetRel )
      I_Contact( #s31_ChkCycleSelect_T1 )
      I_Contact( #s31_ChkCycleSelect_T2 )
      wire#w2
      Coil( #s31_ChkCycleSelect )
   END_RUNG
   RUNG wire#powerrail
      Contact( #s30_WaitCartnSheetOp_T1 )
   END_RUNG wire#w1
   RUNG wire#w2
      { S7_GenerateENO := "TRUE" } Move(in := 31, out1 => #StateNo)
   END_RUNG
   // the same network as SCL:
   #s31_ChkCycleSelect := (#s31_ChkCycleSelect OR #s30_WaitCartnSheetOp_T1) AND NOT #sStWtResetRel AND NOT #s31_ChkCycleSelect_T1 AND NOT #s31_ChkCycleSelect_T2;
   IF #s31_ChkCycleSelect THEN #StateNo := 31; END_IF;
END_REGION

REGION Network 12: Transition for STATE Num:32 Wait for Scan Over
   RUNG wire#powerrail
      Contact( #s32_WaitScanOver )
      I_Contact( #sStWtResetRel )
      Contact( #sSst )
      wire#w1
      Coil( #s32_WaitScanOver_T1 )
   END_RUNG
   RUNG wire#powerrail
      Contact( #iScanOver )
   END_RUNG wire#w1
   RUNG wire#powerrail
      Contact( #iScannerBypass )
   END_RUNG wire#w1
   // the same network as SCL:
   #s32_WaitScanOver_T1 := (#s32_WaitScanOver AND NOT #sStWtResetRel AND #sSst) OR #iScanOver OR #iScannerBypass;
END_REGION

REGION Network 13: STATE Num:32 Wait for Scan Over
   RUNG wire#powerrail
      Contact( #s32_WaitScanOver )
      wire#w1
      I_Contact( #sStWtResetRel )
      I_Contact( #s32_WaitScanOver_T1 )
      wire#w2
      Coil( #s32_WaitScanOver )
   END_RUNG
   RUNG wire#powerrail
      Contact( #s31_ChkCycleSelect_T1 )
   END_RUNG wire#w1
   RUNG wire#w2
      { S7_GenerateENO := "TRUE" } Move(in := 32, out1 => #StateNo)
   END_RUNG
   // the same network as SCL:
   #s32_WaitScanOver := (#s32_WaitScanOver OR #s31_ChkCycleSelect_T1) AND NOT #sStWtResetRel AND NOT #s32_WaitScanOver_T1;
   IF #s32_WaitScanOver THEN #StateNo := 32; END_IF;
END_REGION

REGION Network 14: Actions for STATE Num:32 Wait for Scan Over
   RUNG wire#powerrail
      Contact( #s32_WaitScanOver )
      Coil( #qScanCmd )
   END_RUNG
   // the same network as SCL:
   #qScanCmd := #s32_WaitScanOver;
END_REGION

REGION Network 15: Transition for STATE Num:33 Check Scan result
   RUNG wire#powerrail
      Contact( #s33_ChkScanResult )
      I_Contact( #sStWtResetRel )
      Contact( #sSst )
      wire#w1
      Contact( #iScanOver )
      Contact( #iScanResultOk )
      wire#w2
      Coil( #s33_ChkScanResult_T1 )
   END_RUNG
   RUNG wire#w1
      Contact( #iScannerBypass )
   END_RUNG wire#w2
   RUNG wire#w1
      I_Contact( #s33_ChkScanResult_T1 )
      Contact( #iScanOver )
      Contact( #iScanResultNok )
      Coil( #s33_ChkScanResult_T2 )
   END_RUNG
   // the same network as SCL:
   #_w1 := #s33_ChkScanResult AND NOT #sStWtResetRel AND #sSst;
   #s33_ChkScanResult_T1 := #_w1 AND ((#iScanOver AND #iScanResultOk) OR #iScannerBypass);
   #s33_ChkScanResult_T2 := #_w1 AND NOT #s33_ChkScanResult_T1 AND #iScanOver AND #iScanResultNok;
END_REGION

REGION Network 16: STATE Num:33 Check Scan result
   RUNG wire#powerrail
      Contact( #s33_ChkScanResult )
      wire#w1
      I_Contact( #sStWtResetRel )
      I_Contact( #s33_ChkScanResult_T1 )
      I_Contact( #s33_ChkScanResult_T2 )
      wire#w2
      Coil( #s33_ChkScanResult )
   END_RUNG
   RUNG wire#powerrail
      Contact( #s32_WaitScanOver_T1 )
   END_RUNG wire#w1
   RUNG wire#w2
      { S7_GenerateENO := "TRUE" } Move(in := 33, out1 => #StateNo)
   END_RUNG
   // the same network as SCL:
   #s33_ChkScanResult := (#s33_ChkScanResult OR #s32_WaitScanOver_T1) AND NOT #sStWtResetRel AND NOT #s33_ChkScanResult_T1 AND NOT #s33_ChkScanResult_T2;
   IF #s33_ChkScanResult THEN #StateNo := 33; END_IF;
END_REGION

REGION Network 17: Transition for STATE Num:34 Wait for Operator Decision
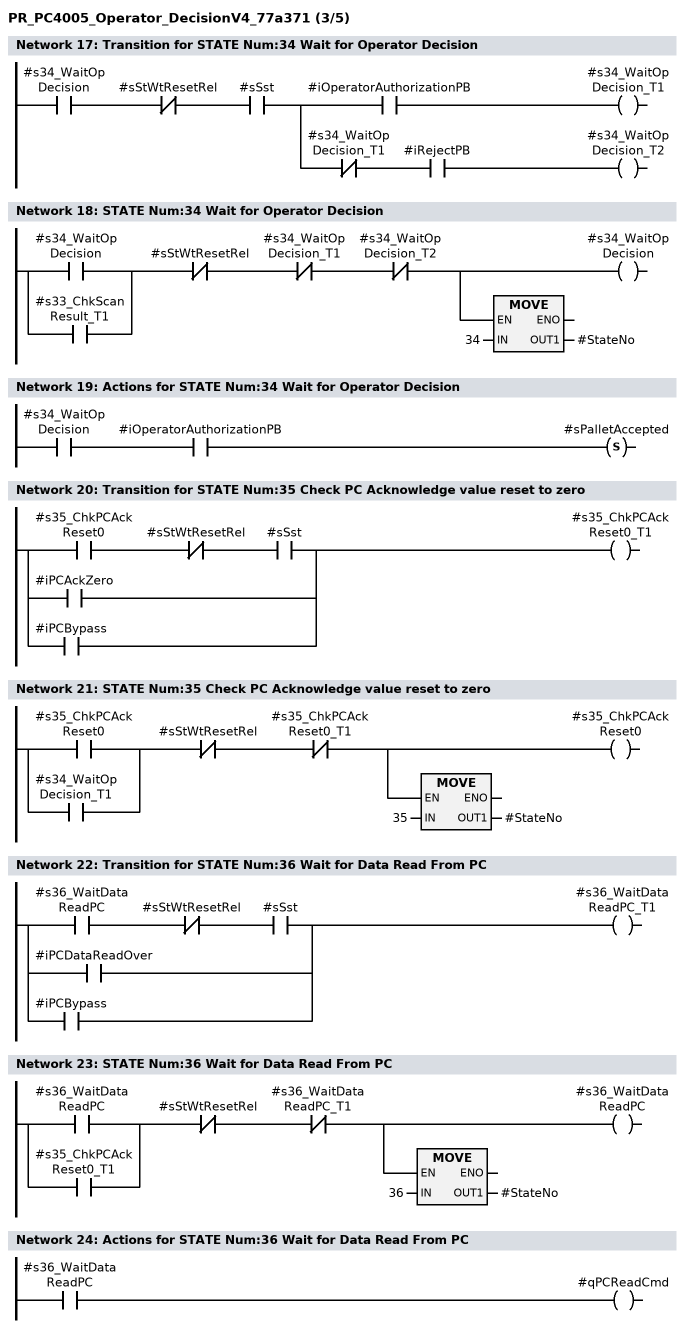
   RUNG wire#powerrail
      Contact( #s34_WaitOpDecision )
      I_Contact( #sStWtResetRel )
      Contact( #sSst )
      wire#w1
      Contact( #iOperatorAuthorizationPB )
      Coil( #s34_WaitOpDecision_T1 )
   END_RUNG
   RUNG wire#w1
      I_Contact( #s34_WaitOpDecision_T1 )
      Contact( #iRejectPB )
      Coil( #s34_WaitOpDecision_T2 )
   END_RUNG
   // the same network as SCL:
   #_w1 := #s34_WaitOpDecision AND NOT #sStWtResetRel AND #sSst;
   #s34_WaitOpDecision_T1 := #_w1 AND #iOperatorAuthorizationPB;
   #s34_WaitOpDecision_T2 := #_w1 AND NOT #s34_WaitOpDecision_T1 AND #iRejectPB;
END_REGION

REGION Network 18: STATE Num:34 Wait for Operator Decision
   RUNG wire#powerrail
      Contact( #s34_WaitOpDecision )
      wire#w1
      I_Contact( #sStWtResetRel )
      I_Contact( #s34_WaitOpDecision_T1 )
      I_Contact( #s34_WaitOpDecision_T2 )
      wire#w2
      Coil( #s34_WaitOpDecision )
   END_RUNG
   RUNG wire#powerrail
      Contact( #s33_ChkScanResult_T1 )
   END_RUNG wire#w1
   RUNG wire#w2
      { S7_GenerateENO := "TRUE" } Move(in := 34, out1 => #StateNo)
   END_RUNG
   // the same network as SCL:
   #s34_WaitOpDecision := (#s34_WaitOpDecision OR #s33_ChkScanResult_T1) AND NOT #sStWtResetRel AND NOT #s34_WaitOpDecision_T1 AND NOT #s34_WaitOpDecision_T2;
   IF #s34_WaitOpDecision THEN #StateNo := 34; END_IF;
END_REGION

REGION Network 19: Actions for STATE Num:34 Wait for Operator Decision
   RUNG wire#powerrail
      Contact( #s34_WaitOpDecision )
      Contact( #iOperatorAuthorizationPB )
      S_Coil( #sPalletAccepted )
   END_RUNG
   // the same network as SCL:
   IF #s34_WaitOpDecision AND #iOperatorAuthorizationPB THEN #sPalletAccepted := TRUE; END_IF;
END_REGION

REGION Network 20: Transition for STATE Num:35 Check PC Acknowledge value reset to zero
   RUNG wire#powerrail
      Contact( #s35_ChkPCAckReset0 )
      I_Contact( #sStWtResetRel )
      Contact( #sSst )
      wire#w1
      Coil( #s35_ChkPCAckReset0_T1 )
   END_RUNG
   RUNG wire#powerrail
      Contact( #iPCAckZero )
   END_RUNG wire#w1
   RUNG wire#powerrail
      Contact( #iPCBypass )
   END_RUNG wire#w1
   // the same network as SCL:
   #s35_ChkPCAckReset0_T1 := (#s35_ChkPCAckReset0 AND NOT #sStWtResetRel AND #sSst) OR #iPCAckZero OR #iPCBypass;
END_REGION

REGION Network 21: STATE Num:35 Check PC Acknowledge value reset to zero
   RUNG wire#powerrail
      Contact( #s35_ChkPCAckReset0 )
      wire#w1
      I_Contact( #sStWtResetRel )
      I_Contact( #s35_ChkPCAckReset0_T1 )
      wire#w2
      Coil( #s35_ChkPCAckReset0 )
   END_RUNG
   RUNG wire#powerrail
      Contact( #s34_WaitOpDecision_T1 )
   END_RUNG wire#w1
   RUNG wire#w2
      { S7_GenerateENO := "TRUE" } Move(in := 35, out1 => #StateNo)
   END_RUNG
   // the same network as SCL:
   #s35_ChkPCAckReset0 := (#s35_ChkPCAckReset0 OR #s34_WaitOpDecision_T1) AND NOT #sStWtResetRel AND NOT #s35_ChkPCAckReset0_T1;
   IF #s35_ChkPCAckReset0 THEN #StateNo := 35; END_IF;
END_REGION

REGION Network 22: Transition for STATE Num:36 Wait for Data Read From PC
   RUNG wire#powerrail
      Contact( #s36_WaitDataReadPC )
      I_Contact( #sStWtResetRel )
      Contact( #sSst )
      wire#w1
      Coil( #s36_WaitDataReadPC_T1 )
   END_RUNG
   RUNG wire#powerrail
      Contact( #iPCDataReadOver )
   END_RUNG wire#w1
   RUNG wire#powerrail
      Contact( #iPCBypass )
   END_RUNG wire#w1
   // the same network as SCL:
   #s36_WaitDataReadPC_T1 := (#s36_WaitDataReadPC AND NOT #sStWtResetRel AND #sSst) OR #iPCDataReadOver OR #iPCBypass;
END_REGION

REGION Network 23: STATE Num:36 Wait for Data Read From PC
   RUNG wire#powerrail
      Contact( #s36_WaitDataReadPC )
      wire#w1
      I_Contact( #sStWtResetRel )
      I_Contact( #s36_WaitDataReadPC_T1 )
      wire#w2
      Coil( #s36_WaitDataReadPC )
   END_RUNG
   RUNG wire#powerrail
      Contact( #s35_ChkPCAckReset0_T1 )
   END_RUNG wire#w1
   RUNG wire#w2
      { S7_GenerateENO := "TRUE" } Move(in := 36, out1 => #StateNo)
   END_RUNG
   // the same network as SCL:
   #s36_WaitDataReadPC := (#s36_WaitDataReadPC OR #s35_ChkPCAckReset0_T1) AND NOT #sStWtResetRel AND NOT #s36_WaitDataReadPC_T1;
   IF #s36_WaitDataReadPC THEN #StateNo := 36; END_IF;
END_REGION

REGION Network 24: Actions for STATE Num:36 Wait for Data Read From PC
   RUNG wire#powerrail
      Contact( #s36_WaitDataReadPC )
      Coil( #qPCReadCmd )
   END_RUNG
   // the same network as SCL:
   #qPCReadCmd := #s36_WaitDataReadPC;
END_REGION

REGION Network 25: Transition for STATE Num:38 Wait for Process Start Low
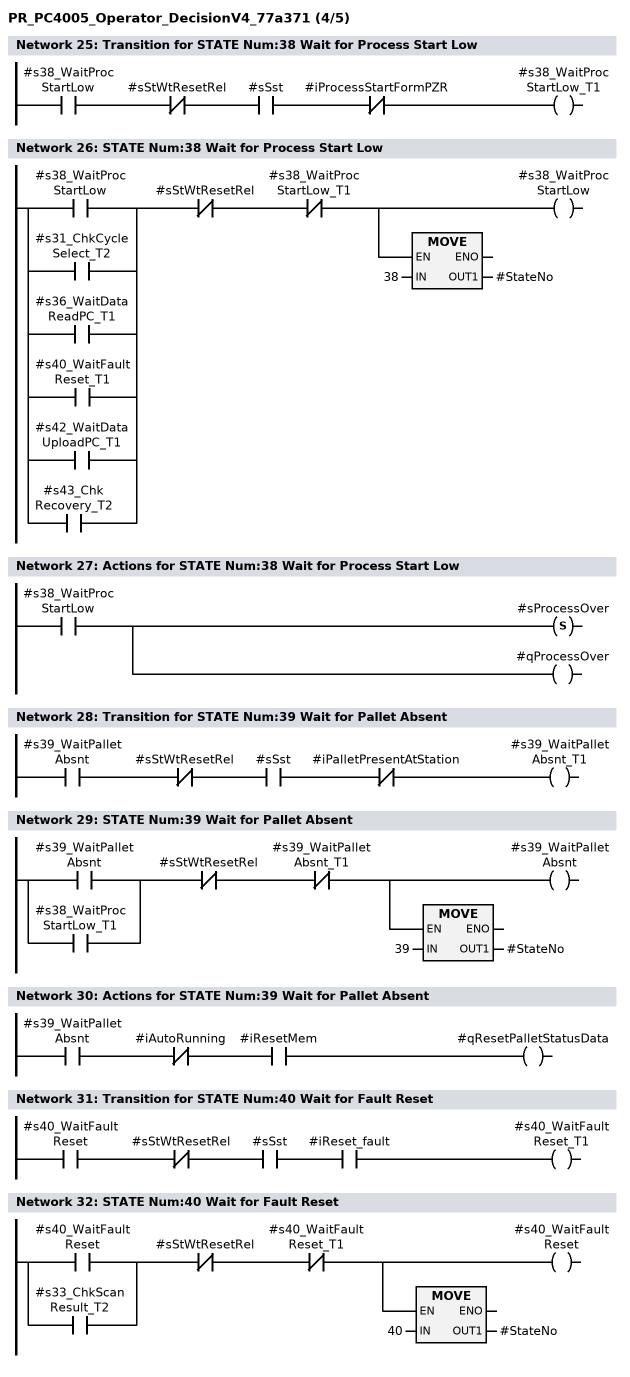
   RUNG wire#powerrail
      Contact( #s38_WaitProcStartLow )
      I_Contact( #sStWtResetRel )
      Contact( #sSst )
      I_Contact( #iProcessStartFormPZR )
      Coil( #s38_WaitProcStartLow_T1 )
   END_RUNG
   // the same network as SCL:
   #s38_WaitProcStartLow_T1 := #s38_WaitProcStartLow AND NOT #sStWtResetRel AND #sSst AND NOT #iProcessStartFormPZR;
END_REGION

REGION Network 26: STATE Num:38 Wait for Process Start Low
   RUNG wire#powerrail
      Contact( #s38_WaitProcStartLow )
      wire#w1
      I_Contact( #sStWtResetRel )
      I_Contact( #s38_WaitProcStartLow_T1 )
      wire#w2
      Coil( #s38_WaitProcStartLow )
   END_RUNG
   RUNG wire#powerrail
      Contact( #s31_ChkCycleSelect_T2 )
   END_RUNG wire#w1
   RUNG wire#powerrail
      Contact( #s36_WaitDataReadPC_T1 )
   END_RUNG wire#w1
   RUNG wire#powerrail
      Contact( #s40_WaitFaultReset_T1 )
   END_RUNG wire#w1
   RUNG wire#powerrail
      Contact( #s42_WaitDataUploadPC_T1 )
   END_RUNG wire#w1
   RUNG wire#powerrail
      Contact( #s43_ChkRecovery_T2 )
   END_RUNG wire#w1
   RUNG wire#w2
      { S7_GenerateENO := "TRUE" } Move(in := 38, out1 => #StateNo)
   END_RUNG
   // the same network as SCL:
   #s38_WaitProcStartLow := (#s38_WaitProcStartLow OR #s31_ChkCycleSelect_T2 OR #s36_WaitDataReadPC_T1 OR #s40_WaitFaultReset_T1 OR #s42_WaitDataUploadPC_T1 OR #s43_ChkRecovery_T2) AND NOT #sStWtResetRel AND NOT #s38_WaitProcStartLow_T1;
   IF #s38_WaitProcStartLow THEN #StateNo := 38; END_IF;
END_REGION

REGION Network 27: Actions for STATE Num:38 Wait for Process Start Low
   RUNG wire#powerrail
      Contact( #s38_WaitProcStartLow )
      wire#w1
      S_Coil( #sProcessOver )
   END_RUNG
   RUNG wire#w1
      Coil( #qProcessOver )
   END_RUNG
   // the same network as SCL:
   IF #s38_WaitProcStartLow THEN #sProcessOver := TRUE; END_IF;
   #qProcessOver := #s38_WaitProcStartLow;
END_REGION

REGION Network 28: Transition for STATE Num:39 Wait for Pallet Absent
   RUNG wire#powerrail
      Contact( #s39_WaitPalletAbsnt )
      I_Contact( #sStWtResetRel )
      Contact( #sSst )
      I_Contact( #iPalletPresentAtStation )
      Coil( #s39_WaitPalletAbsnt_T1 )
   END_RUNG
   // the same network as SCL:
   #s39_WaitPalletAbsnt_T1 := #s39_WaitPalletAbsnt AND NOT #sStWtResetRel AND #sSst AND NOT #iPalletPresentAtStation;
END_REGION

REGION Network 29: STATE Num:39 Wait for Pallet Absent
   RUNG wire#powerrail
      Contact( #s39_WaitPalletAbsnt )
      wire#w1
      I_Contact( #sStWtResetRel )
      I_Contact( #s39_WaitPalletAbsnt_T1 )
      wire#w2
      Coil( #s39_WaitPalletAbsnt )
   END_RUNG
   RUNG wire#powerrail
      Contact( #s38_WaitProcStartLow_T1 )
   END_RUNG wire#w1
   RUNG wire#w2
      { S7_GenerateENO := "TRUE" } Move(in := 39, out1 => #StateNo)
   END_RUNG
   // the same network as SCL:
   #s39_WaitPalletAbsnt := (#s39_WaitPalletAbsnt OR #s38_WaitProcStartLow_T1) AND NOT #sStWtResetRel AND NOT #s39_WaitPalletAbsnt_T1;
   IF #s39_WaitPalletAbsnt THEN #StateNo := 39; END_IF;
END_REGION

REGION Network 30: Actions for STATE Num:39 Wait for Pallet Absent
   RUNG wire#powerrail
      Contact( #s39_WaitPalletAbsnt )
      I_Contact( #iAutoRunning )
      Contact( #iResetMem )
      Coil( #qResetPalletStatusData )
   END_RUNG
   // the same network as SCL:
   #qResetPalletStatusData := #s39_WaitPalletAbsnt AND NOT #iAutoRunning AND #iResetMem;
END_REGION

REGION Network 31: Transition for STATE Num:40 Wait for Fault Reset
   RUNG wire#powerrail
      Contact( #s40_WaitFaultReset )
      I_Contact( #sStWtResetRel )
      Contact( #sSst )
      Contact( #iReset_fault )
      Coil( #s40_WaitFaultReset_T1 )
   END_RUNG
   // the same network as SCL:
   #s40_WaitFaultReset_T1 := #s40_WaitFaultReset AND NOT #sStWtResetRel AND #sSst AND #iReset_fault;
END_REGION

REGION Network 32: STATE Num:40 Wait for Fault Reset
   RUNG wire#powerrail
      Contact( #s40_WaitFaultReset )
      wire#w1
      I_Contact( #sStWtResetRel )
      I_Contact( #s40_WaitFaultReset_T1 )
      wire#w2
      Coil( #s40_WaitFaultReset )
   END_RUNG
   RUNG wire#powerrail
      Contact( #s33_ChkScanResult_T2 )
   END_RUNG wire#w1
   RUNG wire#w2
      { S7_GenerateENO := "TRUE" } Move(in := 40, out1 => #StateNo)
   END_RUNG
   // the same network as SCL:
   #s40_WaitFaultReset := (#s40_WaitFaultReset OR #s33_ChkScanResult_T2) AND NOT #sStWtResetRel AND NOT #s40_WaitFaultReset_T1;
   IF #s40_WaitFaultReset THEN #StateNo := 40; END_IF;
END_REGION

REGION Network 33: Transition for STATE Num:41 Check PC Acknowledge value reset to zero for Upload
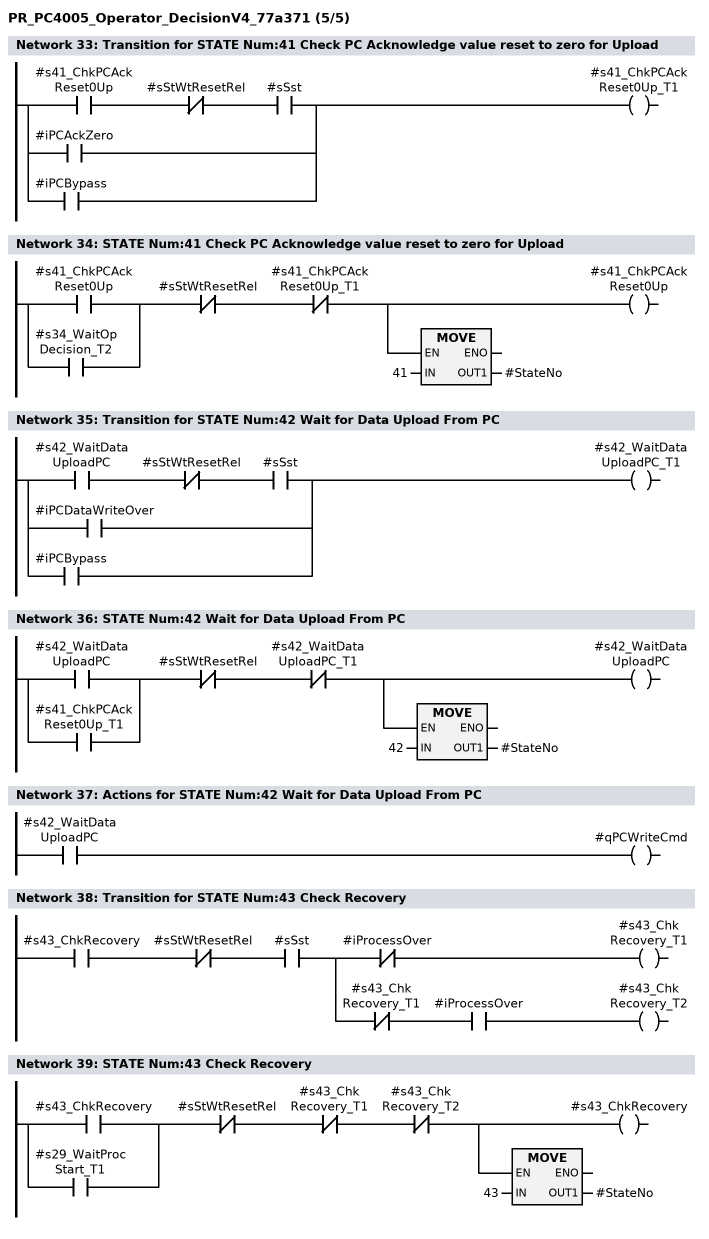
   RUNG wire#powerrail
      Contact( #s41_ChkPCAckReset0Up )
      I_Contact( #sStWtResetRel )
      Contact( #sSst )
      wire#w1
      Coil( #s41_ChkPCAckReset0Up_T1 )
   END_RUNG
   RUNG wire#powerrail
      Contact( #iPCAckZero )
   END_RUNG wire#w1
   RUNG wire#powerrail
      Contact( #iPCBypass )
   END_RUNG wire#w1
   // the same network as SCL:
   #s41_ChkPCAckReset0Up_T1 := (#s41_ChkPCAckReset0Up AND NOT #sStWtResetRel AND #sSst) OR #iPCAckZero OR #iPCBypass;
END_REGION

REGION Network 34: STATE Num:41 Check PC Acknowledge value reset to zero for Upload
   RUNG wire#powerrail
      Contact( #s41_ChkPCAckReset0Up )
      wire#w1
      I_Contact( #sStWtResetRel )
      I_Contact( #s41_ChkPCAckReset0Up_T1 )
      wire#w2
      Coil( #s41_ChkPCAckReset0Up )
   END_RUNG
   RUNG wire#powerrail
      Contact( #s34_WaitOpDecision_T2 )
   END_RUNG wire#w1
   RUNG wire#w2
      { S7_GenerateENO := "TRUE" } Move(in := 41, out1 => #StateNo)
   END_RUNG
   // the same network as SCL:
   #s41_ChkPCAckReset0Up := (#s41_ChkPCAckReset0Up OR #s34_WaitOpDecision_T2) AND NOT #sStWtResetRel AND NOT #s41_ChkPCAckReset0Up_T1;
   IF #s41_ChkPCAckReset0Up THEN #StateNo := 41; END_IF;
END_REGION

REGION Network 35: Transition for STATE Num:42 Wait for Data Upload From PC
   RUNG wire#powerrail
      Contact( #s42_WaitDataUploadPC )
      I_Contact( #sStWtResetRel )
      Contact( #sSst )
      wire#w1
      Coil( #s42_WaitDataUploadPC_T1 )
   END_RUNG
   RUNG wire#powerrail
      Contact( #iPCDataWriteOver )
   END_RUNG wire#w1
   RUNG wire#powerrail
      Contact( #iPCBypass )
   END_RUNG wire#w1
   // the same network as SCL:
   #s42_WaitDataUploadPC_T1 := (#s42_WaitDataUploadPC AND NOT #sStWtResetRel AND #sSst) OR #iPCDataWriteOver OR #iPCBypass;
END_REGION

REGION Network 36: STATE Num:42 Wait for Data Upload From PC
   RUNG wire#powerrail
      Contact( #s42_WaitDataUploadPC )
      wire#w1
      I_Contact( #sStWtResetRel )
      I_Contact( #s42_WaitDataUploadPC_T1 )
      wire#w2
      Coil( #s42_WaitDataUploadPC )
   END_RUNG
   RUNG wire#powerrail
      Contact( #s41_ChkPCAckReset0Up_T1 )
   END_RUNG wire#w1
   RUNG wire#w2
      { S7_GenerateENO := "TRUE" } Move(in := 42, out1 => #StateNo)
   END_RUNG
   // the same network as SCL:
   #s42_WaitDataUploadPC := (#s42_WaitDataUploadPC OR #s41_ChkPCAckReset0Up_T1) AND NOT #sStWtResetRel AND NOT #s42_WaitDataUploadPC_T1;
   IF #s42_WaitDataUploadPC THEN #StateNo := 42; END_IF;
END_REGION

REGION Network 37: Actions for STATE Num:42 Wait for Data Upload From PC
   RUNG wire#powerrail
      Contact( #s42_WaitDataUploadPC )
      Coil( #qPCWriteCmd )
   END_RUNG
   // the same network as SCL:
   #qPCWriteCmd := #s42_WaitDataUploadPC;
END_REGION

REGION Network 38: Transition for STATE Num:43 Check Recovery
   RUNG wire#powerrail
      Contact( #s43_ChkRecovery )
      I_Contact( #sStWtResetRel )
      Contact( #sSst )
      wire#w1
      I_Contact( #iProcessOver )
      Coil( #s43_ChkRecovery_T1 )
   END_RUNG
   RUNG wire#w1
      I_Contact( #s43_ChkRecovery_T1 )
      Contact( #iProcessOver )
      Coil( #s43_ChkRecovery_T2 )
   END_RUNG
   // the same network as SCL:
   #_w1 := #s43_ChkRecovery AND NOT #sStWtResetRel AND #sSst;
   #s43_ChkRecovery_T1 := #_w1 AND NOT #iProcessOver;
   #s43_ChkRecovery_T2 := #_w1 AND NOT #s43_ChkRecovery_T1 AND #iProcessOver;
END_REGION

REGION Network 39: STATE Num:43 Check Recovery
   RUNG wire#powerrail
      Contact( #s43_ChkRecovery )
      wire#w1
      I_Contact( #sStWtResetRel )
      I_Contact( #s43_ChkRecovery_T1 )
      I_Contact( #s43_ChkRecovery_T2 )
      wire#w2
      Coil( #s43_ChkRecovery )
   END_RUNG
   RUNG wire#powerrail
      Contact( #s29_WaitProcStart_T1 )
   END_RUNG wire#w1
   RUNG wire#w2
      { S7_GenerateENO := "TRUE" } Move(in := 43, out1 => #StateNo)
   END_RUNG
   // the same network as SCL:
   #s43_ChkRecovery := (#s43_ChkRecovery OR #s29_WaitProcStart_T1) AND NOT #sStWtResetRel AND NOT #s43_ChkRecovery_T1 AND NOT #s43_ChkRecovery_T2;
   IF #s43_ChkRecovery THEN #StateNo := 43; END_IF;
END_REGION
END_FUNCTION_BLOCK

FUNCTION_BLOCK "PR_PC4005_Operator_DecisionV4_d15416"   // FB2, LAD
VERSION : 0.1
// stored: AutoNumber true, IsIECCheckEnabled false, UDAEnableTagReadback false
   VAR_INPUT
      iAutoRunning : Bool;
      iOperatorAuthorizationPB : Bool;
      iPCAckZero : Bool;
      iPCBypass : Bool;
      iPCDataReadOver : Bool;
      iPCDataWriteOver : Bool;
      iPalletPresentAtStation : Bool;
      iProcessOver : Bool;
      iProcessStartFormPZR : Bool;
      iRejectPB : Bool;
      iResetMem : Bool;
      iReset_fault : Bool;
      iScanOver : Bool;
      iScanResultNok : Bool;
      iScanResultOk : Bool;
      iScannerBypass : Bool;
      iSstMode : Bool;
      iSstPB : Bool;
      iUnloadCycleSelection : Bool;
   END_VAR
   VAR_OUTPUT
      qPCReadCmd : Bool;
      qPCWriteCmd : Bool;
      qProcessOver : Bool;
      qResetPalletStatusData : Bool;
      qScanCmd : Bool;
   END_VAR
   VAR DB_SPECIFIC
      StateNo : Int;
      s29_WaitProcStart : Bool;
      s29_WaitProcStart_T1 : Bool;
      s30_WaitCartnSheetOp : Bool;
      s30_WaitCartnSheetOp_T1 : Bool;
      s31_ChkCycleSelect : Bool;
      s31_ChkCycleSelect_T1 : Bool;
      s31_ChkCycleSelect_T2 : Bool;
      s32_WaitScanOver : Bool;
      s32_WaitScanOver_T1 : Bool;
      s33_ChkScanResult : Bool;
      s33_ChkScanResult_T1 : Bool;
      s33_ChkScanResult_T2 : Bool;
      s34_WaitOpDecision : Bool;
      s34_WaitOpDecision_T1 : Bool;
      s34_WaitOpDecision_T2 : Bool;
      s35_ChkPCAckReset0 : Bool;
      s35_ChkPCAckReset0_T1 : Bool;
      s36_WaitDataReadPC : Bool;
      s36_WaitDataReadPC_T1 : Bool;
      s38_WaitProcStartLow : Bool;
      s38_WaitProcStartLow_T1 : Bool;
      s39_WaitPalletAbsnt : Bool;
      s39_WaitPalletAbsnt_T1 : Bool;
      s40_WaitFaultReset : Bool;
      s40_WaitFaultReset_T1 : Bool;
      s41_ChkPCAckReset0Up : Bool;
      s41_ChkPCAckReset0Up_T1 : Bool;
      s42_WaitDataUploadPC : Bool;
      s42_WaitDataUploadPC_T1 : Bool;
      s43_ChkRecovery : Bool;
      s43_ChkRecovery_T1 : Bool;
      s43_ChkRecovery_T2 : Bool;
      sPalletAccepted : Bool;
      sProcessOver : Bool;
      sSst : Bool;
      sSstPulse : Bool;
      sSstRise : Bool;
      sStWtResetRel : Bool;
      sStWtResetRel_T1 : Bool;
   END_VAR
   VAR_TEMP
      tOne : Bool;
   END_VAR
   VAR_TEMP   // added for the SCL form of the ladder/FBD networks
      _w1 : Bool;
   END_VAR
BEGIN

REGION Network 1
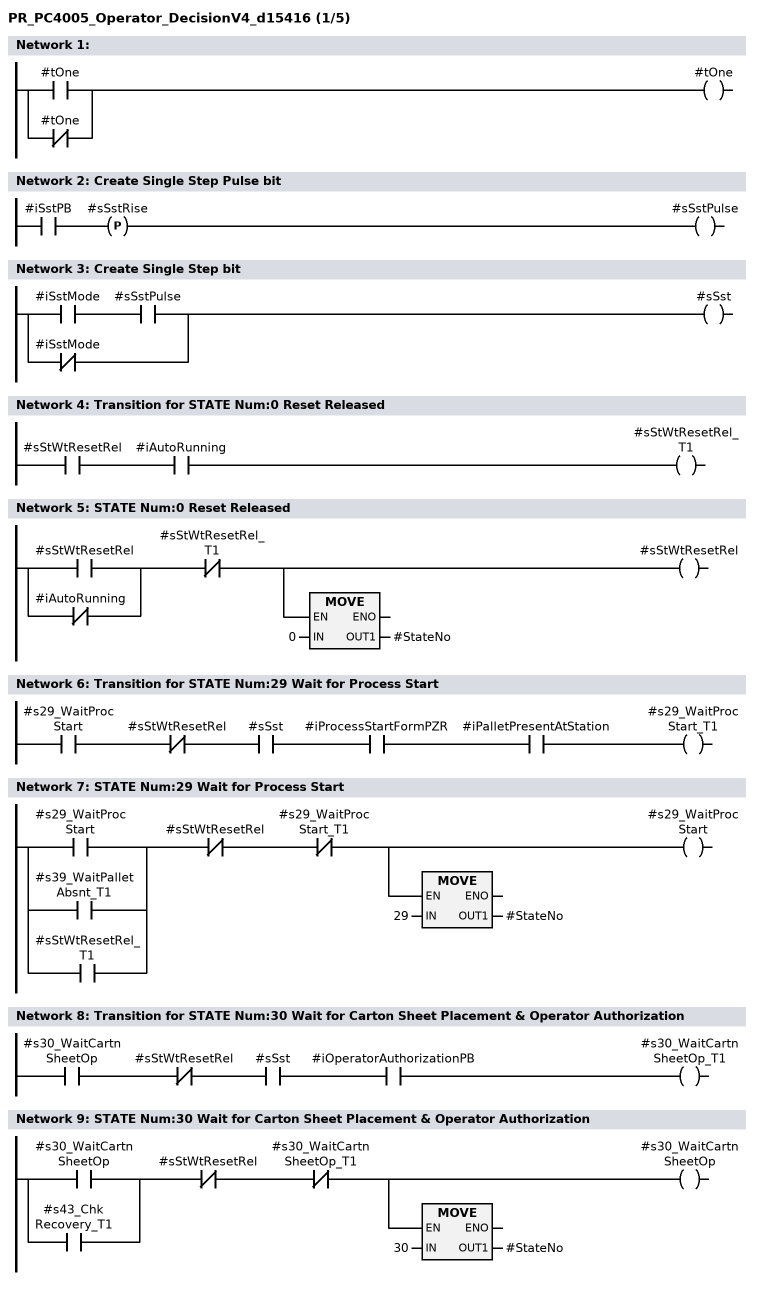
   RUNG wire#powerrail
      Contact( #tOne )
      wire#w1
      Coil( #tOne )
   END_RUNG
   RUNG wire#powerrail
      I_Contact( #tOne )
   END_RUNG wire#w1
   // the same network as SCL:
   #tOne := #tOne OR NOT #tOne;
END_REGION

REGION Network 2: Create Single Step Pulse bit
   RUNG wire#powerrail
      Contact( #iSstPB )
      P_Trig( #sSstRise )
      Coil( #sSstPulse )
   END_RUNG
   // the same network as SCL:
   #_w1 := #iSstPB AND NOT #sSstRise;   // rising edge
   #sSstRise := #iSstPB;
   #sSstPulse := #_w1;
END_REGION

REGION Network 3: Create Single Step bit
   RUNG wire#powerrail
      Contact( #iSstMode )
      Contact( #sSstPulse )
      wire#w1
      Coil( #sSst )
   END_RUNG
   RUNG wire#powerrail
      I_Contact( #iSstMode )
   END_RUNG wire#w1
   // the same network as SCL:
   #sSst := (#iSstMode AND #sSstPulse) OR NOT #iSstMode;
END_REGION

REGION Network 4: Transition for STATE Num:0 Reset Released
   RUNG wire#powerrail
      Contact( #sStWtResetRel )
      Contact( #iAutoRunning )
      Coil( #sStWtResetRel_T1 )
   END_RUNG
   // the same network as SCL:
   #sStWtResetRel_T1 := #sStWtResetRel AND #iAutoRunning;
END_REGION

REGION Network 5: STATE Num:0 Reset Released
   RUNG wire#powerrail
      Contact( #sStWtResetRel )
      wire#w1
      I_Contact( #sStWtResetRel_T1 )
      wire#w2
      Coil( #sStWtResetRel )
   END_RUNG
   RUNG wire#powerrail
      I_Contact( #iAutoRunning )
   END_RUNG wire#w1
   RUNG wire#w2
      { S7_GenerateENO := "TRUE" } Move(in := 0, out1 => #StateNo)
   END_RUNG
   // the same network as SCL:
   #sStWtResetRel := (#sStWtResetRel OR NOT #iAutoRunning) AND NOT #sStWtResetRel_T1;
   IF #sStWtResetRel THEN #StateNo := 0; END_IF;
END_REGION

REGION Network 6: Transition for STATE Num:29 Wait for Process Start
   RUNG wire#powerrail
      Contact( #s29_WaitProcStart )
      I_Contact( #sStWtResetRel )
      Contact( #sSst )
      Contact( #iProcessStartFormPZR )
      Contact( #iPalletPresentAtStation )
      Coil( #s29_WaitProcStart_T1 )
   END_RUNG
   // the same network as SCL:
   #s29_WaitProcStart_T1 := #s29_WaitProcStart AND NOT #sStWtResetRel AND #sSst AND #iProcessStartFormPZR AND #iPalletPresentAtStation;
END_REGION

REGION Network 7: STATE Num:29 Wait for Process Start
   RUNG wire#powerrail
      Contact( #s29_WaitProcStart )
      wire#w1
      I_Contact( #sStWtResetRel )
      I_Contact( #s29_WaitProcStart_T1 )
      wire#w2
      Coil( #s29_WaitProcStart )
   END_RUNG
   RUNG wire#powerrail
      Contact( #s39_WaitPalletAbsnt_T1 )
   END_RUNG wire#w1
   RUNG wire#powerrail
      Contact( #sStWtResetRel_T1 )
   END_RUNG wire#w1
   RUNG wire#w2
      { S7_GenerateENO := "TRUE" } Move(in := 29, out1 => #StateNo)
   END_RUNG
   // the same network as SCL:
   #s29_WaitProcStart := (#s29_WaitProcStart OR #s39_WaitPalletAbsnt_T1 OR #sStWtResetRel_T1) AND NOT #sStWtResetRel AND NOT #s29_WaitProcStart_T1;
   IF #s29_WaitProcStart THEN #StateNo := 29; END_IF;
END_REGION

REGION Network 8: Transition for STATE Num:30 Wait for Carton Sheet Placement & Operator Authorization
   RUNG wire#powerrail
      Contact( #s30_WaitCartnSheetOp )
      I_Contact( #sStWtResetRel )
      Contact( #sSst )
      Contact( #iOperatorAuthorizationPB )
      Coil( #s30_WaitCartnSheetOp_T1 )
   END_RUNG
   // the same network as SCL:
   #s30_WaitCartnSheetOp_T1 := #s30_WaitCartnSheetOp AND NOT #sStWtResetRel AND #sSst AND #iOperatorAuthorizationPB;
END_REGION

REGION Network 9: STATE Num:30 Wait for Carton Sheet Placement & Operator Authorization
   RUNG wire#powerrail
      Contact( #s30_WaitCartnSheetOp )
      wire#w1
      I_Contact( #sStWtResetRel )
      I_Contact( #s30_WaitCartnSheetOp_T1 )
      wire#w2
      Coil( #s30_WaitCartnSheetOp )
   END_RUNG
   RUNG wire#powerrail
      Contact( #s43_ChkRecovery_T1 )
   END_RUNG wire#w1
   RUNG wire#w2
      { S7_GenerateENO := "TRUE" } Move(in := 30, out1 => #StateNo)
   END_RUNG
   // the same network as SCL:
   #s30_WaitCartnSheetOp := (#s30_WaitCartnSheetOp OR #s43_ChkRecovery_T1) AND NOT #sStWtResetRel AND NOT #s30_WaitCartnSheetOp_T1;
   IF #s30_WaitCartnSheetOp THEN #StateNo := 30; END_IF;
END_REGION

REGION Network 10: Transition for STATE Num:31 Check Cycle Selection
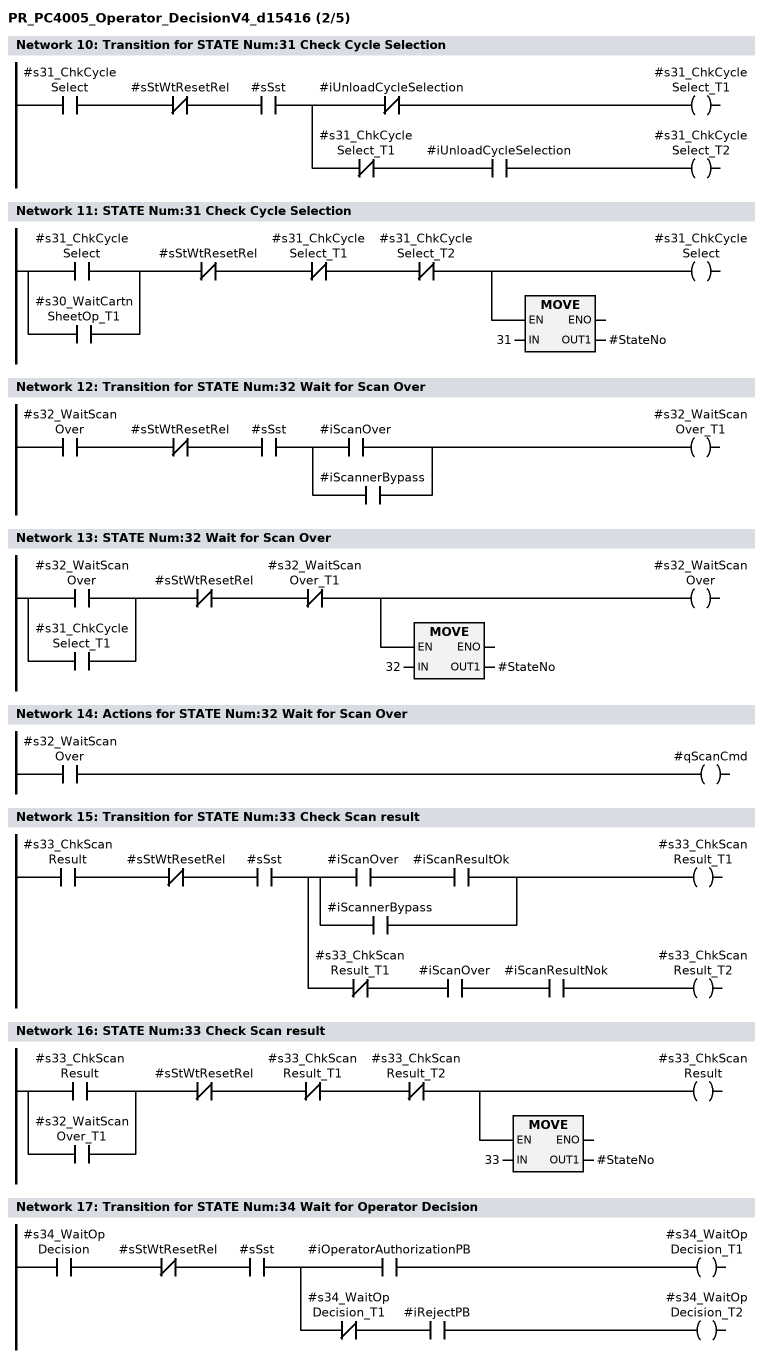
   RUNG wire#powerrail
      Contact( #s31_ChkCycleSelect )
      I_Contact( #sStWtResetRel )
      Contact( #sSst )
      wire#w1
      I_Contact( #iUnloadCycleSelection )
      Coil( #s31_ChkCycleSelect_T1 )
   END_RUNG
   RUNG wire#w1
      I_Contact( #s31_ChkCycleSelect_T1 )
      Contact( #iUnloadCycleSelection )
      Coil( #s31_ChkCycleSelect_T2 )
   END_RUNG
   // the same network as SCL:
   #_w1 := #s31_ChkCycleSelect AND NOT #sStWtResetRel AND #sSst;
   #s31_ChkCycleSelect_T1 := #_w1 AND NOT #iUnloadCycleSelection;
   #s31_ChkCycleSelect_T2 := #_w1 AND NOT #s31_ChkCycleSelect_T1 AND #iUnloadCycleSelection;
END_REGION

REGION Network 11: STATE Num:31 Check Cycle Selection
   RUNG wire#powerrail
      Contact( #s31_ChkCycleSelect )
      wire#w1
      I_Contact( #sStWtResetRel )
      I_Contact( #s31_ChkCycleSelect_T1 )
      I_Contact( #s31_ChkCycleSelect_T2 )
      wire#w2
      Coil( #s31_ChkCycleSelect )
   END_RUNG
   RUNG wire#powerrail
      Contact( #s30_WaitCartnSheetOp_T1 )
   END_RUNG wire#w1
   RUNG wire#w2
      { S7_GenerateENO := "TRUE" } Move(in := 31, out1 => #StateNo)
   END_RUNG
   // the same network as SCL:
   #s31_ChkCycleSelect := (#s31_ChkCycleSelect OR #s30_WaitCartnSheetOp_T1) AND NOT #sStWtResetRel AND NOT #s31_ChkCycleSelect_T1 AND NOT #s31_ChkCycleSelect_T2;
   IF #s31_ChkCycleSelect THEN #StateNo := 31; END_IF;
END_REGION

REGION Network 12: Transition for STATE Num:32 Wait for Scan Over
   RUNG wire#powerrail
      Contact( #s32_WaitScanOver )
      I_Contact( #sStWtResetRel )
      Contact( #sSst )
      wire#w1
      Contact( #iScanOver )
      wire#w2
      Coil( #s32_WaitScanOver_T1 )
   END_RUNG
   RUNG wire#w1
      Contact( #iScannerBypass )
   END_RUNG wire#w2
   // the same network as SCL:
   #s32_WaitScanOver_T1 := #s32_WaitScanOver AND NOT #sStWtResetRel AND #sSst AND (#iScanOver OR #iScannerBypass);
END_REGION

REGION Network 13: STATE Num:32 Wait for Scan Over
   RUNG wire#powerrail
      Contact( #s32_WaitScanOver )
      wire#w1
      I_Contact( #sStWtResetRel )
      I_Contact( #s32_WaitScanOver_T1 )
      wire#w2
      Coil( #s32_WaitScanOver )
   END_RUNG
   RUNG wire#powerrail
      Contact( #s31_ChkCycleSelect_T1 )
   END_RUNG wire#w1
   RUNG wire#w2
      { S7_GenerateENO := "TRUE" } Move(in := 32, out1 => #StateNo)
   END_RUNG
   // the same network as SCL:
   #s32_WaitScanOver := (#s32_WaitScanOver OR #s31_ChkCycleSelect_T1) AND NOT #sStWtResetRel AND NOT #s32_WaitScanOver_T1;
   IF #s32_WaitScanOver THEN #StateNo := 32; END_IF;
END_REGION

REGION Network 14: Actions for STATE Num:32 Wait for Scan Over
   RUNG wire#powerrail
      Contact( #s32_WaitScanOver )
      Coil( #qScanCmd )
   END_RUNG
   // the same network as SCL:
   #qScanCmd := #s32_WaitScanOver;
END_REGION

REGION Network 15: Transition for STATE Num:33 Check Scan result
   RUNG wire#powerrail
      Contact( #s33_ChkScanResult )
      I_Contact( #sStWtResetRel )
      Contact( #sSst )
      wire#w1
      Contact( #iScanOver )
      Contact( #iScanResultOk )
      wire#w2
      Coil( #s33_ChkScanResult_T1 )
   END_RUNG
   RUNG wire#w1
      Contact( #iScannerBypass )
   END_RUNG wire#w2
   RUNG wire#w1
      I_Contact( #s33_ChkScanResult_T1 )
      Contact( #iScanOver )
      Contact( #iScanResultNok )
      Coil( #s33_ChkScanResult_T2 )
   END_RUNG
   // the same network as SCL:
   #_w1 := #s33_ChkScanResult AND NOT #sStWtResetRel AND #sSst;
   #s33_ChkScanResult_T1 := #_w1 AND ((#iScanOver AND #iScanResultOk) OR #iScannerBypass);
   #s33_ChkScanResult_T2 := #_w1 AND NOT #s33_ChkScanResult_T1 AND #iScanOver AND #iScanResultNok;
END_REGION

REGION Network 16: STATE Num:33 Check Scan result
   RUNG wire#powerrail
      Contact( #s33_ChkScanResult )
      wire#w1
      I_Contact( #sStWtResetRel )
      I_Contact( #s33_ChkScanResult_T1 )
      I_Contact( #s33_ChkScanResult_T2 )
      wire#w2
      Coil( #s33_ChkScanResult )
   END_RUNG
   RUNG wire#powerrail
      Contact( #s32_WaitScanOver_T1 )
   END_RUNG wire#w1
   RUNG wire#w2
      { S7_GenerateENO := "TRUE" } Move(in := 33, out1 => #StateNo)
   END_RUNG
   // the same network as SCL:
   #s33_ChkScanResult := (#s33_ChkScanResult OR #s32_WaitScanOver_T1) AND NOT #sStWtResetRel AND NOT #s33_ChkScanResult_T1 AND NOT #s33_ChkScanResult_T2;
   IF #s33_ChkScanResult THEN #StateNo := 33; END_IF;
END_REGION

REGION Network 17: Transition for STATE Num:34 Wait for Operator Decision
   RUNG wire#powerrail
      Contact( #s34_WaitOpDecision )
      I_Contact( #sStWtResetRel )
      Contact( #sSst )
      wire#w1
      Contact( #iOperatorAuthorizationPB )
      Coil( #s34_WaitOpDecision_T1 )
   END_RUNG
   RUNG wire#w1
      I_Contact( #s34_WaitOpDecision_T1 )
      Contact( #iRejectPB )
      Coil( #s34_WaitOpDecision_T2 )
   END_RUNG
   // the same network as SCL:
   #_w1 := #s34_WaitOpDecision AND NOT #sStWtResetRel AND #sSst;
   #s34_WaitOpDecision_T1 := #_w1 AND #iOperatorAuthorizationPB;
   #s34_WaitOpDecision_T2 := #_w1 AND NOT #s34_WaitOpDecision_T1 AND #iRejectPB;
END_REGION

REGION Network 18: STATE Num:34 Wait for Operator Decision
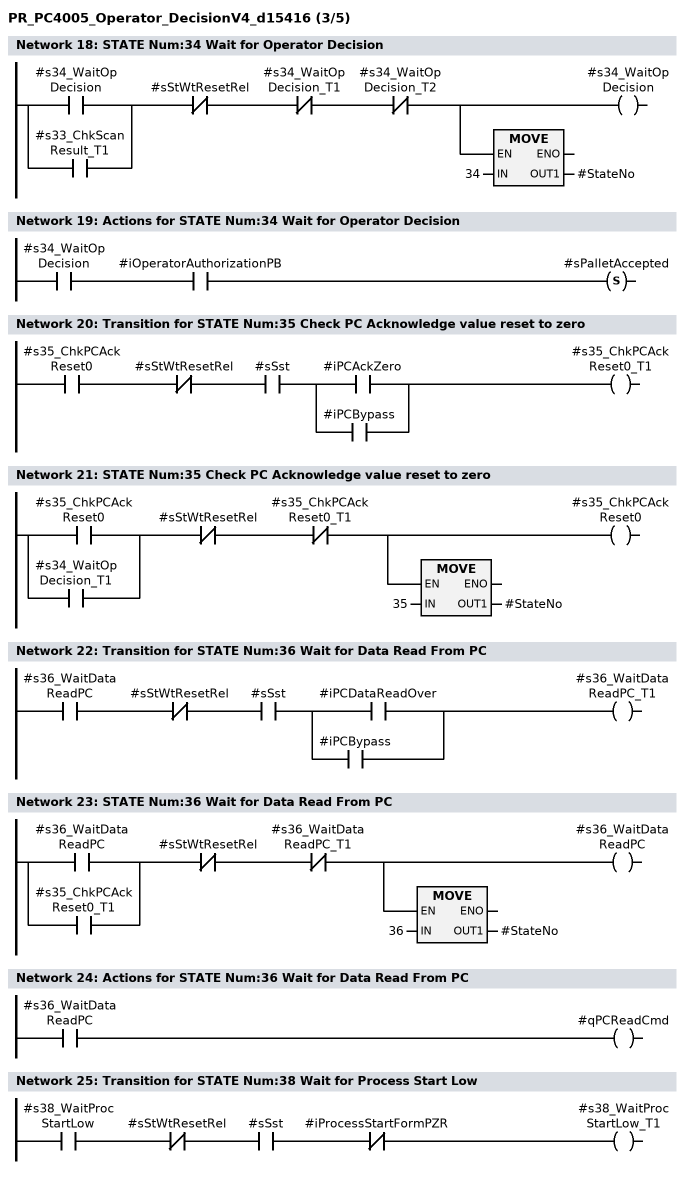
   RUNG wire#powerrail
      Contact( #s34_WaitOpDecision )
      wire#w1
      I_Contact( #sStWtResetRel )
      I_Contact( #s34_WaitOpDecision_T1 )
      I_Contact( #s34_WaitOpDecision_T2 )
      wire#w2
      Coil( #s34_WaitOpDecision )
   END_RUNG
   RUNG wire#powerrail
      Contact( #s33_ChkScanResult_T1 )
   END_RUNG wire#w1
   RUNG wire#w2
      { S7_GenerateENO := "TRUE" } Move(in := 34, out1 => #StateNo)
   END_RUNG
   // the same network as SCL:
   #s34_WaitOpDecision := (#s34_WaitOpDecision OR #s33_ChkScanResult_T1) AND NOT #sStWtResetRel AND NOT #s34_WaitOpDecision_T1 AND NOT #s34_WaitOpDecision_T2;
   IF #s34_WaitOpDecision THEN #StateNo := 34; END_IF;
END_REGION

REGION Network 19: Actions for STATE Num:34 Wait for Operator Decision
   RUNG wire#powerrail
      Contact( #s34_WaitOpDecision )
      Contact( #iOperatorAuthorizationPB )
      S_Coil( #sPalletAccepted )
   END_RUNG
   // the same network as SCL:
   IF #s34_WaitOpDecision AND #iOperatorAuthorizationPB THEN #sPalletAccepted := TRUE; END_IF;
END_REGION

REGION Network 20: Transition for STATE Num:35 Check PC Acknowledge value reset to zero
   RUNG wire#powerrail
      Contact( #s35_ChkPCAckReset0 )
      I_Contact( #sStWtResetRel )
      Contact( #sSst )
      wire#w1
      Contact( #iPCAckZero )
      wire#w2
      Coil( #s35_ChkPCAckReset0_T1 )
   END_RUNG
   RUNG wire#w1
      Contact( #iPCBypass )
   END_RUNG wire#w2
   // the same network as SCL:
   #s35_ChkPCAckReset0_T1 := #s35_ChkPCAckReset0 AND NOT #sStWtResetRel AND #sSst AND (#iPCAckZero OR #iPCBypass);
END_REGION

REGION Network 21: STATE Num:35 Check PC Acknowledge value reset to zero
   RUNG wire#powerrail
      Contact( #s35_ChkPCAckReset0 )
      wire#w1
      I_Contact( #sStWtResetRel )
      I_Contact( #s35_ChkPCAckReset0_T1 )
      wire#w2
      Coil( #s35_ChkPCAckReset0 )
   END_RUNG
   RUNG wire#powerrail
      Contact( #s34_WaitOpDecision_T1 )
   END_RUNG wire#w1
   RUNG wire#w2
      { S7_GenerateENO := "TRUE" } Move(in := 35, out1 => #StateNo)
   END_RUNG
   // the same network as SCL:
   #s35_ChkPCAckReset0 := (#s35_ChkPCAckReset0 OR #s34_WaitOpDecision_T1) AND NOT #sStWtResetRel AND NOT #s35_ChkPCAckReset0_T1;
   IF #s35_ChkPCAckReset0 THEN #StateNo := 35; END_IF;
END_REGION

REGION Network 22: Transition for STATE Num:36 Wait for Data Read From PC
   RUNG wire#powerrail
      Contact( #s36_WaitDataReadPC )
      I_Contact( #sStWtResetRel )
      Contact( #sSst )
      wire#w1
      Contact( #iPCDataReadOver )
      wire#w2
      Coil( #s36_WaitDataReadPC_T1 )
   END_RUNG
   RUNG wire#w1
      Contact( #iPCBypass )
   END_RUNG wire#w2
   // the same network as SCL:
   #s36_WaitDataReadPC_T1 := #s36_WaitDataReadPC AND NOT #sStWtResetRel AND #sSst AND (#iPCDataReadOver OR #iPCBypass);
END_REGION

REGION Network 23: STATE Num:36 Wait for Data Read From PC
   RUNG wire#powerrail
      Contact( #s36_WaitDataReadPC )
      wire#w1
      I_Contact( #sStWtResetRel )
      I_Contact( #s36_WaitDataReadPC_T1 )
      wire#w2
      Coil( #s36_WaitDataReadPC )
   END_RUNG
   RUNG wire#powerrail
      Contact( #s35_ChkPCAckReset0_T1 )
   END_RUNG wire#w1
   RUNG wire#w2
      { S7_GenerateENO := "TRUE" } Move(in := 36, out1 => #StateNo)
   END_RUNG
   // the same network as SCL:
   #s36_WaitDataReadPC := (#s36_WaitDataReadPC OR #s35_ChkPCAckReset0_T1) AND NOT #sStWtResetRel AND NOT #s36_WaitDataReadPC_T1;
   IF #s36_WaitDataReadPC THEN #StateNo := 36; END_IF;
END_REGION

REGION Network 24: Actions for STATE Num:36 Wait for Data Read From PC
   RUNG wire#powerrail
      Contact( #s36_WaitDataReadPC )
      Coil( #qPCReadCmd )
   END_RUNG
   // the same network as SCL:
   #qPCReadCmd := #s36_WaitDataReadPC;
END_REGION

REGION Network 25: Transition for STATE Num:38 Wait for Process Start Low
   RUNG wire#powerrail
      Contact( #s38_WaitProcStartLow )
      I_Contact( #sStWtResetRel )
      Contact( #sSst )
      I_Contact( #iProcessStartFormPZR )
      Coil( #s38_WaitProcStartLow_T1 )
   END_RUNG
   // the same network as SCL:
   #s38_WaitProcStartLow_T1 := #s38_WaitProcStartLow AND NOT #sStWtResetRel AND #sSst AND NOT #iProcessStartFormPZR;
END_REGION

REGION Network 26: STATE Num:38 Wait for Process Start Low
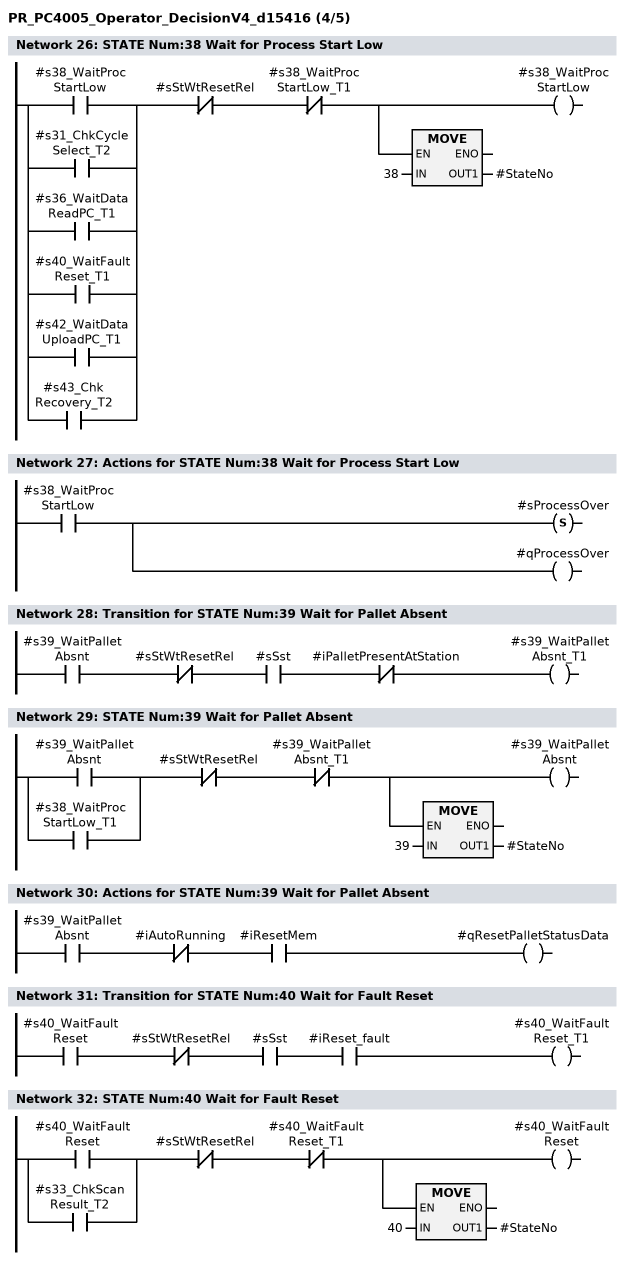
   RUNG wire#powerrail
      Contact( #s38_WaitProcStartLow )
      wire#w1
      I_Contact( #sStWtResetRel )
      I_Contact( #s38_WaitProcStartLow_T1 )
      wire#w2
      Coil( #s38_WaitProcStartLow )
   END_RUNG
   RUNG wire#powerrail
      Contact( #s31_ChkCycleSelect_T2 )
   END_RUNG wire#w1
   RUNG wire#powerrail
      Contact( #s36_WaitDataReadPC_T1 )
   END_RUNG wire#w1
   RUNG wire#powerrail
      Contact( #s40_WaitFaultReset_T1 )
   END_RUNG wire#w1
   RUNG wire#powerrail
      Contact( #s42_WaitDataUploadPC_T1 )
   END_RUNG wire#w1
   RUNG wire#powerrail
      Contact( #s43_ChkRecovery_T2 )
   END_RUNG wire#w1
   RUNG wire#w2
      { S7_GenerateENO := "TRUE" } Move(in := 38, out1 => #StateNo)
   END_RUNG
   // the same network as SCL:
   #s38_WaitProcStartLow := (#s38_WaitProcStartLow OR #s31_ChkCycleSelect_T2 OR #s36_WaitDataReadPC_T1 OR #s40_WaitFaultReset_T1 OR #s42_WaitDataUploadPC_T1 OR #s43_ChkRecovery_T2) AND NOT #sStWtResetRel AND NOT #s38_WaitProcStartLow_T1;
   IF #s38_WaitProcStartLow THEN #StateNo := 38; END_IF;
END_REGION

REGION Network 27: Actions for STATE Num:38 Wait for Process Start Low
   RUNG wire#powerrail
      Contact( #s38_WaitProcStartLow )
      wire#w1
      S_Coil( #sProcessOver )
   END_RUNG
   RUNG wire#w1
      Coil( #qProcessOver )
   END_RUNG
   // the same network as SCL:
   IF #s38_WaitProcStartLow THEN #sProcessOver := TRUE; END_IF;
   #qProcessOver := #s38_WaitProcStartLow;
END_REGION

REGION Network 28: Transition for STATE Num:39 Wait for Pallet Absent
   RUNG wire#powerrail
      Contact( #s39_WaitPalletAbsnt )
      I_Contact( #sStWtResetRel )
      Contact( #sSst )
      I_Contact( #iPalletPresentAtStation )
      Coil( #s39_WaitPalletAbsnt_T1 )
   END_RUNG
   // the same network as SCL:
   #s39_WaitPalletAbsnt_T1 := #s39_WaitPalletAbsnt AND NOT #sStWtResetRel AND #sSst AND NOT #iPalletPresentAtStation;
END_REGION

REGION Network 29: STATE Num:39 Wait for Pallet Absent
   RUNG wire#powerrail
      Contact( #s39_WaitPalletAbsnt )
      wire#w1
      I_Contact( #sStWtResetRel )
      I_Contact( #s39_WaitPalletAbsnt_T1 )
      wire#w2
      Coil( #s39_WaitPalletAbsnt )
   END_RUNG
   RUNG wire#powerrail
      Contact( #s38_WaitProcStartLow_T1 )
   END_RUNG wire#w1
   RUNG wire#w2
      { S7_GenerateENO := "TRUE" } Move(in := 39, out1 => #StateNo)
   END_RUNG
   // the same network as SCL:
   #s39_WaitPalletAbsnt := (#s39_WaitPalletAbsnt OR #s38_WaitProcStartLow_T1) AND NOT #sStWtResetRel AND NOT #s39_WaitPalletAbsnt_T1;
   IF #s39_WaitPalletAbsnt THEN #StateNo := 39; END_IF;
END_REGION

REGION Network 30: Actions for STATE Num:39 Wait for Pallet Absent
   RUNG wire#powerrail
      Contact( #s39_WaitPalletAbsnt )
      I_Contact( #iAutoRunning )
      Contact( #iResetMem )
      Coil( #qResetPalletStatusData )
   END_RUNG
   // the same network as SCL:
   #qResetPalletStatusData := #s39_WaitPalletAbsnt AND NOT #iAutoRunning AND #iResetMem;
END_REGION

REGION Network 31: Transition for STATE Num:40 Wait for Fault Reset
   RUNG wire#powerrail
      Contact( #s40_WaitFaultReset )
      I_Contact( #sStWtResetRel )
      Contact( #sSst )
      Contact( #iReset_fault )
      Coil( #s40_WaitFaultReset_T1 )
   END_RUNG
   // the same network as SCL:
   #s40_WaitFaultReset_T1 := #s40_WaitFaultReset AND NOT #sStWtResetRel AND #sSst AND #iReset_fault;
END_REGION

REGION Network 32: STATE Num:40 Wait for Fault Reset
   RUNG wire#powerrail
      Contact( #s40_WaitFaultReset )
      wire#w1
      I_Contact( #sStWtResetRel )
      I_Contact( #s40_WaitFaultReset_T1 )
      wire#w2
      Coil( #s40_WaitFaultReset )
   END_RUNG
   RUNG wire#powerrail
      Contact( #s33_ChkScanResult_T2 )
   END_RUNG wire#w1
   RUNG wire#w2
      { S7_GenerateENO := "TRUE" } Move(in := 40, out1 => #StateNo)
   END_RUNG
   // the same network as SCL:
   #s40_WaitFaultReset := (#s40_WaitFaultReset OR #s33_ChkScanResult_T2) AND NOT #sStWtResetRel AND NOT #s40_WaitFaultReset_T1;
   IF #s40_WaitFaultReset THEN #StateNo := 40; END_IF;
END_REGION

REGION Network 33: Transition for STATE Num:41 Check PC Acknowledge value reset to zero for Upload
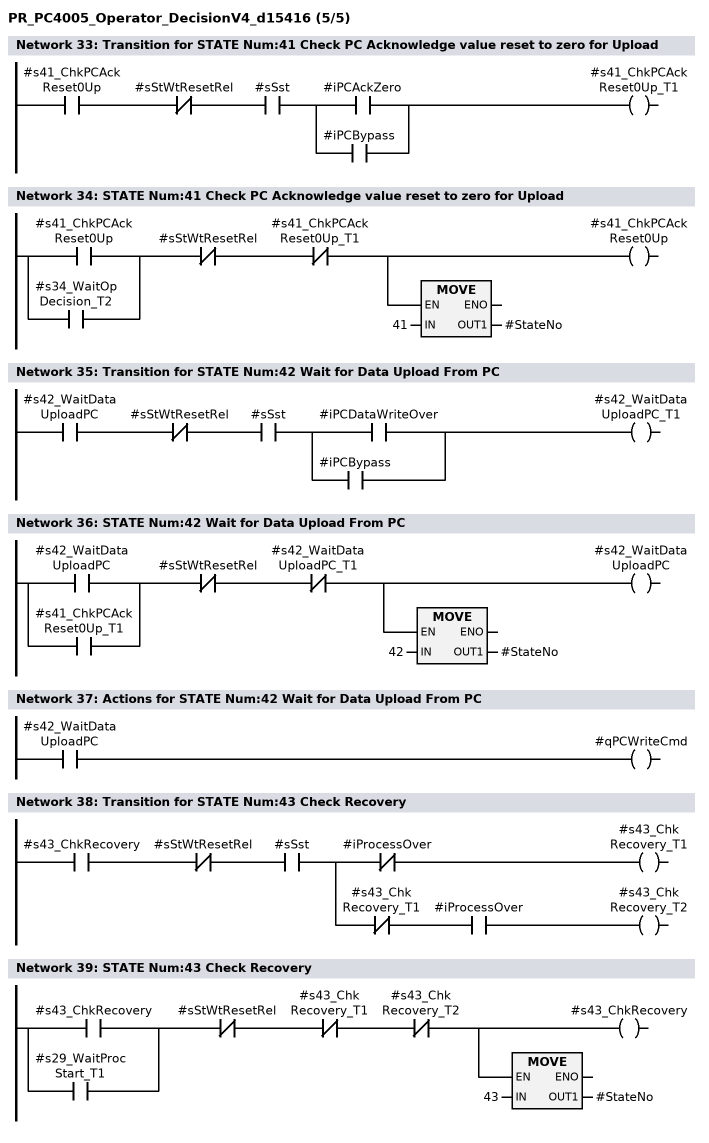
   RUNG wire#powerrail
      Contact( #s41_ChkPCAckReset0Up )
      I_Contact( #sStWtResetRel )
      Contact( #sSst )
      wire#w1
      Contact( #iPCAckZero )
      wire#w2
      Coil( #s41_ChkPCAckReset0Up_T1 )
   END_RUNG
   RUNG wire#w1
      Contact( #iPCBypass )
   END_RUNG wire#w2
   // the same network as SCL:
   #s41_ChkPCAckReset0Up_T1 := #s41_ChkPCAckReset0Up AND NOT #sStWtResetRel AND #sSst AND (#iPCAckZero OR #iPCBypass);
END_REGION

REGION Network 34: STATE Num:41 Check PC Acknowledge value reset to zero for Upload
   RUNG wire#powerrail
      Contact( #s41_ChkPCAckReset0Up )
      wire#w1
      I_Contact( #sStWtResetRel )
      I_Contact( #s41_ChkPCAckReset0Up_T1 )
      wire#w2
      Coil( #s41_ChkPCAckReset0Up )
   END_RUNG
   RUNG wire#powerrail
      Contact( #s34_WaitOpDecision_T2 )
   END_RUNG wire#w1
   RUNG wire#w2
      { S7_GenerateENO := "TRUE" } Move(in := 41, out1 => #StateNo)
   END_RUNG
   // the same network as SCL:
   #s41_ChkPCAckReset0Up := (#s41_ChkPCAckReset0Up OR #s34_WaitOpDecision_T2) AND NOT #sStWtResetRel AND NOT #s41_ChkPCAckReset0Up_T1;
   IF #s41_ChkPCAckReset0Up THEN #StateNo := 41; END_IF;
END_REGION

REGION Network 35: Transition for STATE Num:42 Wait for Data Upload From PC
   RUNG wire#powerrail
      Contact( #s42_WaitDataUploadPC )
      I_Contact( #sStWtResetRel )
      Contact( #sSst )
      wire#w1
      Contact( #iPCDataWriteOver )
      wire#w2
      Coil( #s42_WaitDataUploadPC_T1 )
   END_RUNG
   RUNG wire#w1
      Contact( #iPCBypass )
   END_RUNG wire#w2
   // the same network as SCL:
   #s42_WaitDataUploadPC_T1 := #s42_WaitDataUploadPC AND NOT #sStWtResetRel AND #sSst AND (#iPCDataWriteOver OR #iPCBypass);
END_REGION

REGION Network 36: STATE Num:42 Wait for Data Upload From PC
   RUNG wire#powerrail
      Contact( #s42_WaitDataUploadPC )
      wire#w1
      I_Contact( #sStWtResetRel )
      I_Contact( #s42_WaitDataUploadPC_T1 )
      wire#w2
      Coil( #s42_WaitDataUploadPC )
   END_RUNG
   RUNG wire#powerrail
      Contact( #s41_ChkPCAckReset0Up_T1 )
   END_RUNG wire#w1
   RUNG wire#w2
      { S7_GenerateENO := "TRUE" } Move(in := 42, out1 => #StateNo)
   END_RUNG
   // the same network as SCL:
   #s42_WaitDataUploadPC := (#s42_WaitDataUploadPC OR #s41_ChkPCAckReset0Up_T1) AND NOT #sStWtResetRel AND NOT #s42_WaitDataUploadPC_T1;
   IF #s42_WaitDataUploadPC THEN #StateNo := 42; END_IF;
END_REGION

REGION Network 37: Actions for STATE Num:42 Wait for Data Upload From PC
   RUNG wire#powerrail
      Contact( #s42_WaitDataUploadPC )
      Coil( #qPCWriteCmd )
   END_RUNG
   // the same network as SCL:
   #qPCWriteCmd := #s42_WaitDataUploadPC;
END_REGION

REGION Network 38: Transition for STATE Num:43 Check Recovery
   RUNG wire#powerrail
      Contact( #s43_ChkRecovery )
      I_Contact( #sStWtResetRel )
      Contact( #sSst )
      wire#w1
      I_Contact( #iProcessOver )
      Coil( #s43_ChkRecovery_T1 )
   END_RUNG
   RUNG wire#w1
      I_Contact( #s43_ChkRecovery_T1 )
      Contact( #iProcessOver )
      Coil( #s43_ChkRecovery_T2 )
   END_RUNG
   // the same network as SCL:
   #_w1 := #s43_ChkRecovery AND NOT #sStWtResetRel AND #sSst;
   #s43_ChkRecovery_T1 := #_w1 AND NOT #iProcessOver;
   #s43_ChkRecovery_T2 := #_w1 AND NOT #s43_ChkRecovery_T1 AND #iProcessOver;
END_REGION

REGION Network 39: STATE Num:43 Check Recovery
   RUNG wire#powerrail
      Contact( #s43_ChkRecovery )
      wire#w1
      I_Contact( #sStWtResetRel )
      I_Contact( #s43_ChkRecovery_T1 )
      I_Contact( #s43_ChkRecovery_T2 )
      wire#w2
      Coil( #s43_ChkRecovery )
   END_RUNG
   RUNG wire#powerrail
      Contact( #s29_WaitProcStart_T1 )
   END_RUNG wire#w1
   RUNG wire#w2
      { S7_GenerateENO := "TRUE" } Move(in := 43, out1 => #StateNo)
   END_RUNG
   // the same network as SCL:
   #s43_ChkRecovery := (#s43_ChkRecovery OR #s29_WaitProcStart_T1) AND NOT #sStWtResetRel AND NOT #s43_ChkRecovery_T1 AND NOT #s43_ChkRecovery_T2;
   IF #s43_ChkRecovery THEN #StateNo := 43; END_IF;
END_REGION
END_FUNCTION_BLOCK

FUNCTION_BLOCK "RD_PR_CentreStand_Fix_Seq_V12"   // FB1, LAD
VERSION : 0.1
// stored: AutoNumber true, IsIECCheckEnabled false, UDAEnableTagReadback false
   VAR_INPUT
      iAutoRunning : Bool;
      iFixClamp : Bool;
      iFixEmpty : Bool;
      iFixTrayPresent : Bool;
      iFixUnclamp : Bool;
      iR1DropOver : Bool;
      iR1PickOver : Bool;
      iR2OperationOver : Bool;
      iR2ServiceActivated : Bool;
      iReset_fault : Bool;
      iRobotOutofZone : Bool;
      iSstMode : Bool;
      iSstPB : Bool;
   END_VAR
   VAR_OUTPUT
      qFixClamp : Bool;
      qFixUnclamp : Bool;
      qR1ReadytoDropTray : Bool;
      qR1ReadytoPickTray : Bool;
      qR2OperationStart : Bool;
   END_VAR
   VAR_IN_OUT
      iqR2ServiceActive : Bool;
      iqR2ServiceCompleted : Bool;
   END_VAR
   VAR DB_SPECIFIC
      StateNo : Int;
      s138_WaitBothRbtOutAl : Bool;
      s138_WaitBothRbtOutAl_T1 : Bool;
      s138_WaitBothRbtOutAl_T2 : Bool;
      s139_FixEmpty : Bool;
      s139_FixEmpty_T1 : Bool;
      s140_FixTrayPrsntRec : Bool;
      s140_FixTrayPrsntRec_T1 : Bool;
      s140_FixTrayPrsntRec_T2 : Bool;
      s141_FixUnclampCmd : Bool;
      s141_FixUnclampCmd_T1 : Bool;
      s142_TrayRdyDropFix : Bool;
      s142_TrayRdyDropFix_T1 : Bool;
      s143_RbtDropFixChkTr : Bool;
      s143_RbtDropFixChkTr_T1 : Bool;
      s144_RbtOutAreaDrop : Bool;
      s144_RbtOutAreaDrop_T1 : Bool;
      s145_FixClamp : Bool;
      s145_FixClamp_T1 : Bool;
      s146_Rbt2AlloyOpOver : Bool;
      s146_Rbt2AlloyOpOver_T1 : Bool;
      s147_FixUnclmpCmdAft : Bool;
      s147_FixUnclmpCmdAft_T1 : Bool;
      s148_RdyPickTrayAftr : Bool;
      s148_RdyPickTrayAftr_T1 : Bool;
      s149_RbtPickTrayChkE : Bool;
      s149_RbtPickTrayChkE_T1 : Bool;
      s191_WaitRbt2OutArea : Bool;
      s191_WaitRbt2OutArea_T1 : Bool;
      sSst : Bool;
      sSstPulse : Bool;
      sSstRise : Bool;
      sStWtResetRel : Bool;
      sStWtResetRel_T1 : Bool;
   END_VAR
   VAR_TEMP
      c138_WaitBothRbtOutAl_T1 : Bool;
      c138_WaitBothRbtOutAl_T2 : Bool;
      c140_FixTrayPrsntRec_T1 : Bool;
      c140_FixTrayPrsntRec_T2 : Bool;
      tOne : Bool;
   END_VAR
   VAR_TEMP   // added for the SCL form of the ladder/FBD networks
      _w1 : Bool;
   END_VAR
BEGIN

REGION Network 1
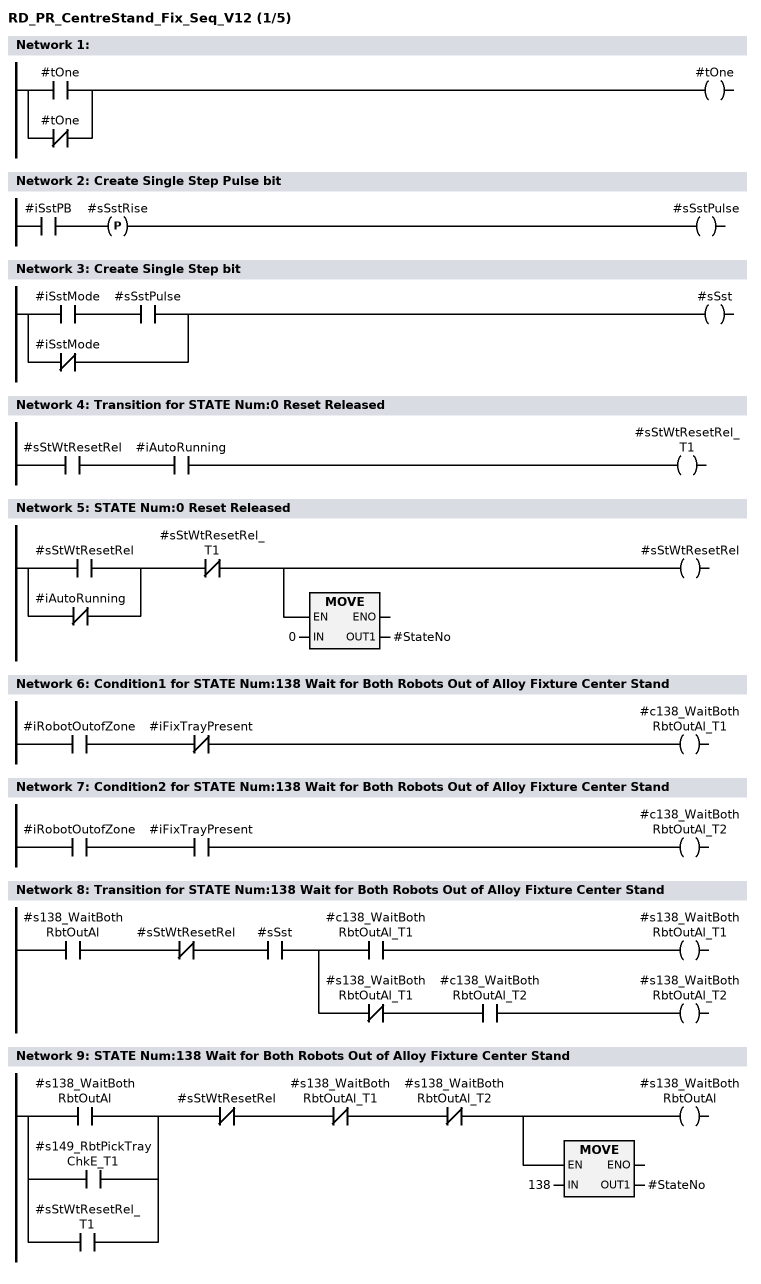
   RUNG wire#powerrail
      Contact( #tOne )
      wire#w1
      Coil( #tOne )
   END_RUNG
   RUNG wire#powerrail
      I_Contact( #tOne )
   END_RUNG wire#w1
   // the same network as SCL:
   #tOne := #tOne OR NOT #tOne;
END_REGION

REGION Network 2: Create Single Step Pulse bit
   RUNG wire#powerrail
      Contact( #iSstPB )
      P_Trig( #sSstRise )
      Coil( #sSstPulse )
   END_RUNG
   // the same network as SCL:
   #_w1 := #iSstPB AND NOT #sSstRise;   // rising edge
   #sSstRise := #iSstPB;
   #sSstPulse := #_w1;
END_REGION

REGION Network 3: Create Single Step bit
   RUNG wire#powerrail
      Contact( #iSstMode )
      Contact( #sSstPulse )
      wire#w1
      Coil( #sSst )
   END_RUNG
   RUNG wire#powerrail
      I_Contact( #iSstMode )
   END_RUNG wire#w1
   // the same network as SCL:
   #sSst := (#iSstMode AND #sSstPulse) OR NOT #iSstMode;
END_REGION

REGION Network 4: Transition for STATE Num:0 Reset Released
   RUNG wire#powerrail
      Contact( #sStWtResetRel )
      Contact( #iAutoRunning )
      Coil( #sStWtResetRel_T1 )
   END_RUNG
   // the same network as SCL:
   #sStWtResetRel_T1 := #sStWtResetRel AND #iAutoRunning;
END_REGION

REGION Network 5: STATE Num:0 Reset Released
   RUNG wire#powerrail
      Contact( #sStWtResetRel )
      wire#w1
      I_Contact( #sStWtResetRel_T1 )
      wire#w2
      Coil( #sStWtResetRel )
   END_RUNG
   RUNG wire#powerrail
      I_Contact( #iAutoRunning )
   END_RUNG wire#w1
   RUNG wire#w2
      { S7_GenerateENO := "TRUE" } Move(in := 0, out1 => #StateNo)
   END_RUNG
   // the same network as SCL:
   #sStWtResetRel := (#sStWtResetRel OR NOT #iAutoRunning) AND NOT #sStWtResetRel_T1;
   IF #sStWtResetRel THEN #StateNo := 0; END_IF;
END_REGION

REGION Network 6: Condition1 for STATE Num:138 Wait for Both Robots Out of Alloy Fixture Center Stand
   RUNG wire#powerrail
      Contact( #iRobotOutofZone )
      I_Contact( #iFixTrayPresent )
      Coil( #c138_WaitBothRbtOutAl_T1 )
   END_RUNG
   // the same network as SCL:
   #c138_WaitBothRbtOutAl_T1 := #iRobotOutofZone AND NOT #iFixTrayPresent;
END_REGION

REGION Network 7: Condition2 for STATE Num:138 Wait for Both Robots Out of Alloy Fixture Center Stand
   RUNG wire#powerrail
      Contact( #iRobotOutofZone )
      Contact( #iFixTrayPresent )
      Coil( #c138_WaitBothRbtOutAl_T2 )
   END_RUNG
   // the same network as SCL:
   #c138_WaitBothRbtOutAl_T2 := #iRobotOutofZone AND #iFixTrayPresent;
END_REGION

REGION Network 8: Transition for STATE Num:138 Wait for Both Robots Out of Alloy Fixture Center Stand
   RUNG wire#powerrail
      Contact( #s138_WaitBothRbtOutAl )
      I_Contact( #sStWtResetRel )
      Contact( #sSst )
      wire#w1
      Contact( #c138_WaitBothRbtOutAl_T1 )
      Coil( #s138_WaitBothRbtOutAl_T1 )
   END_RUNG
   RUNG wire#w1
      I_Contact( #s138_WaitBothRbtOutAl_T1 )
      Contact( #c138_WaitBothRbtOutAl_T2 )
      Coil( #s138_WaitBothRbtOutAl_T2 )
   END_RUNG
   // the same network as SCL:
   #_w1 := #s138_WaitBothRbtOutAl AND NOT #sStWtResetRel AND #sSst;
   #s138_WaitBothRbtOutAl_T1 := #_w1 AND #c138_WaitBothRbtOutAl_T1;
   #s138_WaitBothRbtOutAl_T2 := #_w1 AND NOT #s138_WaitBothRbtOutAl_T1 AND #c138_WaitBothRbtOutAl_T2;
END_REGION

REGION Network 9: STATE Num:138 Wait for Both Robots Out of Alloy Fixture Center Stand
   RUNG wire#powerrail
      Contact( #s138_WaitBothRbtOutAl )
      wire#w1
      I_Contact( #sStWtResetRel )
      I_Contact( #s138_WaitBothRbtOutAl_T1 )
      I_Contact( #s138_WaitBothRbtOutAl_T2 )
      wire#w2
      Coil( #s138_WaitBothRbtOutAl )
   END_RUNG
   RUNG wire#powerrail
      Contact( #s149_RbtPickTrayChkE_T1 )
   END_RUNG wire#w1
   RUNG wire#powerrail
      Contact( #sStWtResetRel_T1 )
   END_RUNG wire#w1
   RUNG wire#w2
      { S7_GenerateENO := "TRUE" } Move(in := 138, out1 => #StateNo)
   END_RUNG
   // the same network as SCL:
   #s138_WaitBothRbtOutAl := (#s138_WaitBothRbtOutAl OR #s149_RbtPickTrayChkE_T1 OR #sStWtResetRel_T1) AND NOT #sStWtResetRel AND NOT #s138_WaitBothRbtOutAl_T1 AND NOT #s138_WaitBothRbtOutAl_T2;
   IF #s138_WaitBothRbtOutAl THEN #StateNo := 138; END_IF;
END_REGION

REGION Network 10: Transition for STATE Num:139 Fix Empty
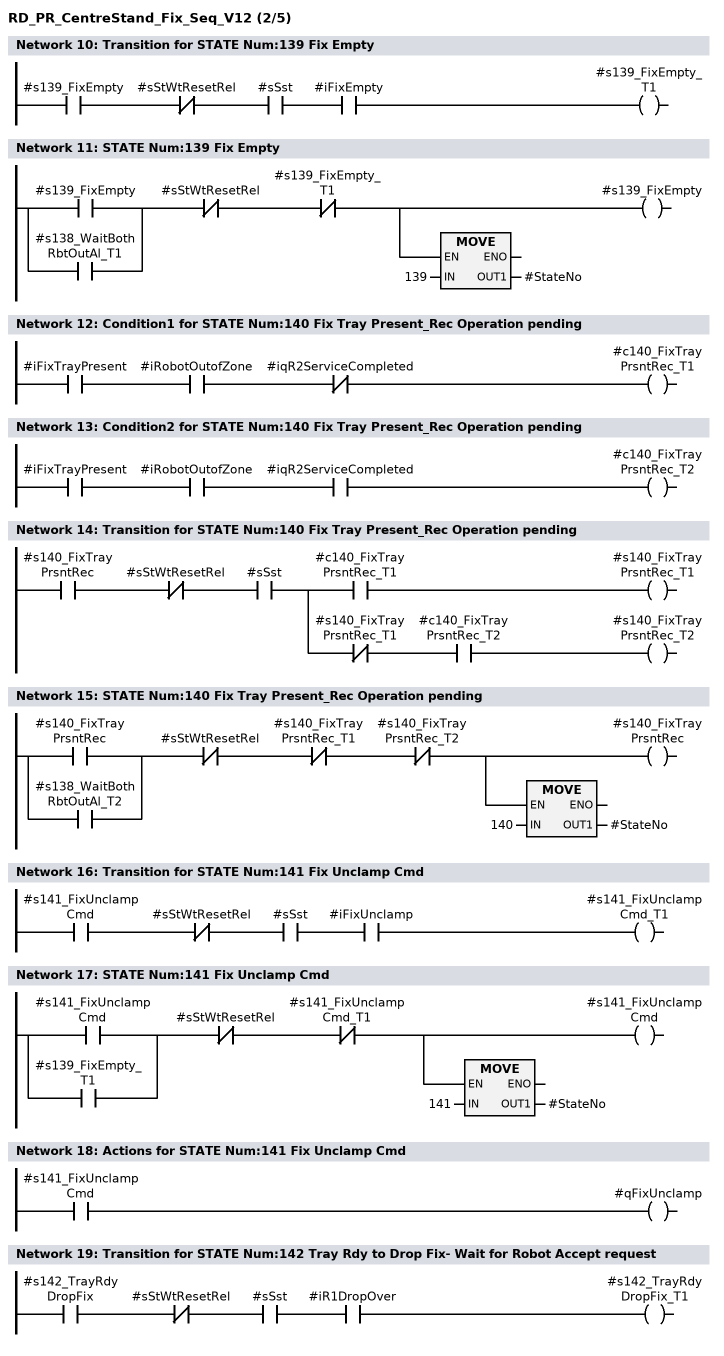
   RUNG wire#powerrail
      Contact( #s139_FixEmpty )
      I_Contact( #sStWtResetRel )
      Contact( #sSst )
      Contact( #iFixEmpty )
      Coil( #s139_FixEmpty_T1 )
   END_RUNG
   // the same network as SCL:
   #s139_FixEmpty_T1 := #s139_FixEmpty AND NOT #sStWtResetRel AND #sSst AND #iFixEmpty;
END_REGION

REGION Network 11: STATE Num:139 Fix Empty
   RUNG wire#powerrail
      Contact( #s139_FixEmpty )
      wire#w1
      I_Contact( #sStWtResetRel )
      I_Contact( #s139_FixEmpty_T1 )
      wire#w2
      Coil( #s139_FixEmpty )
   END_RUNG
   RUNG wire#powerrail
      Contact( #s138_WaitBothRbtOutAl_T1 )
   END_RUNG wire#w1
   RUNG wire#w2
      { S7_GenerateENO := "TRUE" } Move(in := 139, out1 => #StateNo)
   END_RUNG
   // the same network as SCL:
   #s139_FixEmpty := (#s139_FixEmpty OR #s138_WaitBothRbtOutAl_T1) AND NOT #sStWtResetRel AND NOT #s139_FixEmpty_T1;
   IF #s139_FixEmpty THEN #StateNo := 139; END_IF;
END_REGION

REGION Network 12: Condition1 for STATE Num:140 Fix Tray Present_Rec Operation pending
   RUNG wire#powerrail
      Contact( #iFixTrayPresent )
      Contact( #iRobotOutofZone )
      I_Contact( #iqR2ServiceCompleted )
      Coil( #c140_FixTrayPrsntRec_T1 )
   END_RUNG
   // the same network as SCL:
   #c140_FixTrayPrsntRec_T1 := #iFixTrayPresent AND #iRobotOutofZone AND NOT #iqR2ServiceCompleted;
END_REGION

REGION Network 13: Condition2 for STATE Num:140 Fix Tray Present_Rec Operation pending
   RUNG wire#powerrail
      Contact( #iFixTrayPresent )
      Contact( #iRobotOutofZone )
      Contact( #iqR2ServiceCompleted )
      Coil( #c140_FixTrayPrsntRec_T2 )
   END_RUNG
   // the same network as SCL:
   #c140_FixTrayPrsntRec_T2 := #iFixTrayPresent AND #iRobotOutofZone AND #iqR2ServiceCompleted;
END_REGION

REGION Network 14: Transition for STATE Num:140 Fix Tray Present_Rec Operation pending
   RUNG wire#powerrail
      Contact( #s140_FixTrayPrsntRec )
      I_Contact( #sStWtResetRel )
      Contact( #sSst )
      wire#w1
      Contact( #c140_FixTrayPrsntRec_T1 )
      Coil( #s140_FixTrayPrsntRec_T1 )
   END_RUNG
   RUNG wire#w1
      I_Contact( #s140_FixTrayPrsntRec_T1 )
      Contact( #c140_FixTrayPrsntRec_T2 )
      Coil( #s140_FixTrayPrsntRec_T2 )
   END_RUNG
   // the same network as SCL:
   #_w1 := #s140_FixTrayPrsntRec AND NOT #sStWtResetRel AND #sSst;
   #s140_FixTrayPrsntRec_T1 := #_w1 AND #c140_FixTrayPrsntRec_T1;
   #s140_FixTrayPrsntRec_T2 := #_w1 AND NOT #s140_FixTrayPrsntRec_T1 AND #c140_FixTrayPrsntRec_T2;
END_REGION

REGION Network 15: STATE Num:140 Fix Tray Present_Rec Operation pending
   RUNG wire#powerrail
      Contact( #s140_FixTrayPrsntRec )
      wire#w1
      I_Contact( #sStWtResetRel )
      I_Contact( #s140_FixTrayPrsntRec_T1 )
      I_Contact( #s140_FixTrayPrsntRec_T2 )
      wire#w2
      Coil( #s140_FixTrayPrsntRec )
   END_RUNG
   RUNG wire#powerrail
      Contact( #s138_WaitBothRbtOutAl_T2 )
   END_RUNG wire#w1
   RUNG wire#w2
      { S7_GenerateENO := "TRUE" } Move(in := 140, out1 => #StateNo)
   END_RUNG
   // the same network as SCL:
   #s140_FixTrayPrsntRec := (#s140_FixTrayPrsntRec OR #s138_WaitBothRbtOutAl_T2) AND NOT #sStWtResetRel AND NOT #s140_FixTrayPrsntRec_T1 AND NOT #s140_FixTrayPrsntRec_T2;
   IF #s140_FixTrayPrsntRec THEN #StateNo := 140; END_IF;
END_REGION

REGION Network 16: Transition for STATE Num:141 Fix Unclamp Cmd
   RUNG wire#powerrail
      Contact( #s141_FixUnclampCmd )
      I_Contact( #sStWtResetRel )
      Contact( #sSst )
      Contact( #iFixUnclamp )
      Coil( #s141_FixUnclampCmd_T1 )
   END_RUNG
   // the same network as SCL:
   #s141_FixUnclampCmd_T1 := #s141_FixUnclampCmd AND NOT #sStWtResetRel AND #sSst AND #iFixUnclamp;
END_REGION

REGION Network 17: STATE Num:141 Fix Unclamp Cmd
   RUNG wire#powerrail
      Contact( #s141_FixUnclampCmd )
      wire#w1
      I_Contact( #sStWtResetRel )
      I_Contact( #s141_FixUnclampCmd_T1 )
      wire#w2
      Coil( #s141_FixUnclampCmd )
   END_RUNG
   RUNG wire#powerrail
      Contact( #s139_FixEmpty_T1 )
   END_RUNG wire#w1
   RUNG wire#w2
      { S7_GenerateENO := "TRUE" } Move(in := 141, out1 => #StateNo)
   END_RUNG
   // the same network as SCL:
   #s141_FixUnclampCmd := (#s141_FixUnclampCmd OR #s139_FixEmpty_T1) AND NOT #sStWtResetRel AND NOT #s141_FixUnclampCmd_T1;
   IF #s141_FixUnclampCmd THEN #StateNo := 141; END_IF;
END_REGION

REGION Network 18: Actions for STATE Num:141 Fix Unclamp Cmd
   RUNG wire#powerrail
      Contact( #s141_FixUnclampCmd )
      Coil( #qFixUnclamp )
   END_RUNG
   // the same network as SCL:
   #qFixUnclamp := #s141_FixUnclampCmd;
END_REGION

REGION Network 19: Transition for STATE Num:142 Tray Rdy to Drop Fix- Wait for Robot Accept request
   RUNG wire#powerrail
      Contact( #s142_TrayRdyDropFix )
      I_Contact( #sStWtResetRel )
      Contact( #sSst )
      Contact( #iR1DropOver )
      Coil( #s142_TrayRdyDropFix_T1 )
   END_RUNG
   // the same network as SCL:
   #s142_TrayRdyDropFix_T1 := #s142_TrayRdyDropFix AND NOT #sStWtResetRel AND #sSst AND #iR1DropOver;
END_REGION

REGION Network 20: STATE Num:142 Tray Rdy to Drop Fix- Wait for Robot Accept request
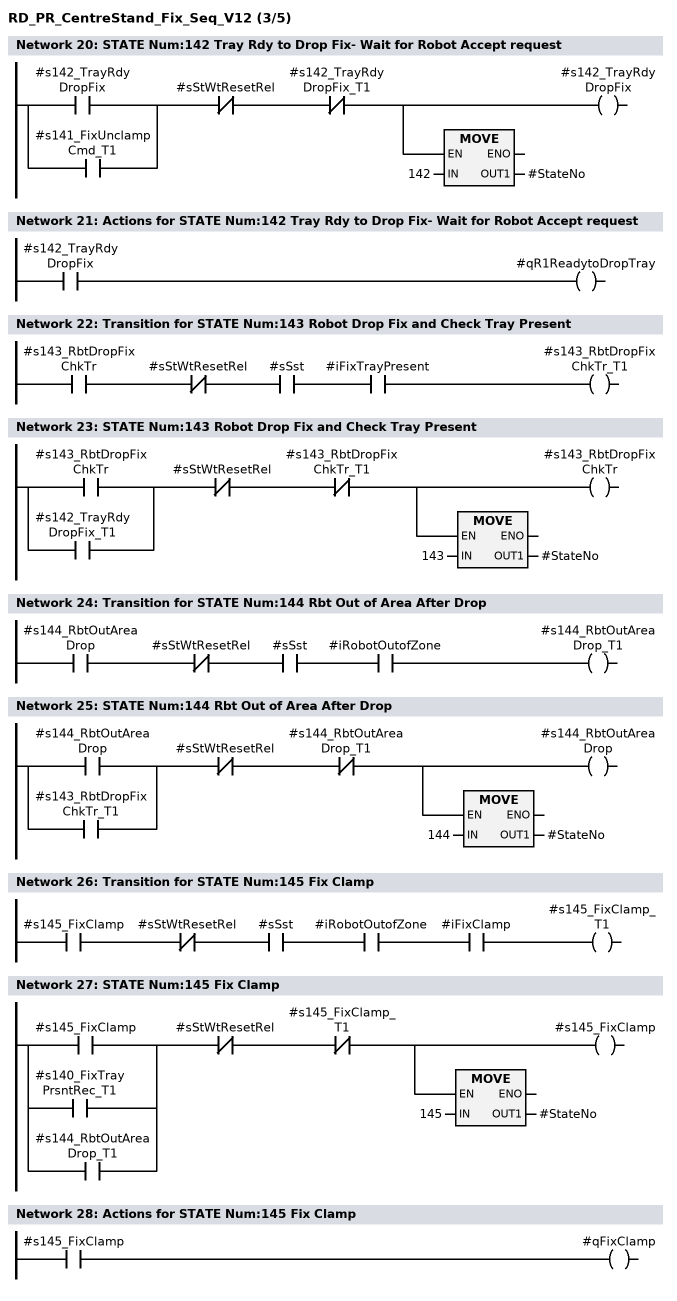
   RUNG wire#powerrail
      Contact( #s142_TrayRdyDropFix )
      wire#w1
      I_Contact( #sStWtResetRel )
      I_Contact( #s142_TrayRdyDropFix_T1 )
      wire#w2
      Coil( #s142_TrayRdyDropFix )
   END_RUNG
   RUNG wire#powerrail
      Contact( #s141_FixUnclampCmd_T1 )
   END_RUNG wire#w1
   RUNG wire#w2
      { S7_GenerateENO := "TRUE" } Move(in := 142, out1 => #StateNo)
   END_RUNG
   // the same network as SCL:
   #s142_TrayRdyDropFix := (#s142_TrayRdyDropFix OR #s141_FixUnclampCmd_T1) AND NOT #sStWtResetRel AND NOT #s142_TrayRdyDropFix_T1;
   IF #s142_TrayRdyDropFix THEN #StateNo := 142; END_IF;
END_REGION

REGION Network 21: Actions for STATE Num:142 Tray Rdy to Drop Fix- Wait for Robot Accept request
   RUNG wire#powerrail
      Contact( #s142_TrayRdyDropFix )
      Coil( #qR1ReadytoDropTray )
   END_RUNG
   // the same network as SCL:
   #qR1ReadytoDropTray := #s142_TrayRdyDropFix;
END_REGION

REGION Network 22: Transition for STATE Num:143 Robot Drop Fix and Check Tray Present
   RUNG wire#powerrail
      Contact( #s143_RbtDropFixChkTr )
      I_Contact( #sStWtResetRel )
      Contact( #sSst )
      Contact( #iFixTrayPresent )
      Coil( #s143_RbtDropFixChkTr_T1 )
   END_RUNG
   // the same network as SCL:
   #s143_RbtDropFixChkTr_T1 := #s143_RbtDropFixChkTr AND NOT #sStWtResetRel AND #sSst AND #iFixTrayPresent;
END_REGION

REGION Network 23: STATE Num:143 Robot Drop Fix and Check Tray Present
   RUNG wire#powerrail
      Contact( #s143_RbtDropFixChkTr )
      wire#w1
      I_Contact( #sStWtResetRel )
      I_Contact( #s143_RbtDropFixChkTr_T1 )
      wire#w2
      Coil( #s143_RbtDropFixChkTr )
   END_RUNG
   RUNG wire#powerrail
      Contact( #s142_TrayRdyDropFix_T1 )
   END_RUNG wire#w1
   RUNG wire#w2
      { S7_GenerateENO := "TRUE" } Move(in := 143, out1 => #StateNo)
   END_RUNG
   // the same network as SCL:
   #s143_RbtDropFixChkTr := (#s143_RbtDropFixChkTr OR #s142_TrayRdyDropFix_T1) AND NOT #sStWtResetRel AND NOT #s143_RbtDropFixChkTr_T1;
   IF #s143_RbtDropFixChkTr THEN #StateNo := 143; END_IF;
END_REGION

REGION Network 24: Transition for STATE Num:144 Rbt Out of Area After Drop
   RUNG wire#powerrail
      Contact( #s144_RbtOutAreaDrop )
      I_Contact( #sStWtResetRel )
      Contact( #sSst )
      Contact( #iRobotOutofZone )
      Coil( #s144_RbtOutAreaDrop_T1 )
   END_RUNG
   // the same network as SCL:
   #s144_RbtOutAreaDrop_T1 := #s144_RbtOutAreaDrop AND NOT #sStWtResetRel AND #sSst AND #iRobotOutofZone;
END_REGION

REGION Network 25: STATE Num:144 Rbt Out of Area After Drop
   RUNG wire#powerrail
      Contact( #s144_RbtOutAreaDrop )
      wire#w1
      I_Contact( #sStWtResetRel )
      I_Contact( #s144_RbtOutAreaDrop_T1 )
      wire#w2
      Coil( #s144_RbtOutAreaDrop )
   END_RUNG
   RUNG wire#powerrail
      Contact( #s143_RbtDropFixChkTr_T1 )
   END_RUNG wire#w1
   RUNG wire#w2
      { S7_GenerateENO := "TRUE" } Move(in := 144, out1 => #StateNo)
   END_RUNG
   // the same network as SCL:
   #s144_RbtOutAreaDrop := (#s144_RbtOutAreaDrop OR #s143_RbtDropFixChkTr_T1) AND NOT #sStWtResetRel AND NOT #s144_RbtOutAreaDrop_T1;
   IF #s144_RbtOutAreaDrop THEN #StateNo := 144; END_IF;
END_REGION

REGION Network 26: Transition for STATE Num:145 Fix Clamp
   RUNG wire#powerrail
      Contact( #s145_FixClamp )
      I_Contact( #sStWtResetRel )
      Contact( #sSst )
      Contact( #iRobotOutofZone )
      Contact( #iFixClamp )
      Coil( #s145_FixClamp_T1 )
   END_RUNG
   // the same network as SCL:
   #s145_FixClamp_T1 := #s145_FixClamp AND NOT #sStWtResetRel AND #sSst AND #iRobotOutofZone AND #iFixClamp;
END_REGION

REGION Network 27: STATE Num:145 Fix Clamp
   RUNG wire#powerrail
      Contact( #s145_FixClamp )
      wire#w1
      I_Contact( #sStWtResetRel )
      I_Contact( #s145_FixClamp_T1 )
      wire#w2
      Coil( #s145_FixClamp )
   END_RUNG
   RUNG wire#powerrail
      Contact( #s140_FixTrayPrsntRec_T1 )
   END_RUNG wire#w1
   RUNG wire#powerrail
      Contact( #s144_RbtOutAreaDrop_T1 )
   END_RUNG wire#w1
   RUNG wire#w2
      { S7_GenerateENO := "TRUE" } Move(in := 145, out1 => #StateNo)
   END_RUNG
   // the same network as SCL:
   #s145_FixClamp := (#s145_FixClamp OR #s140_FixTrayPrsntRec_T1 OR #s144_RbtOutAreaDrop_T1) AND NOT #sStWtResetRel AND NOT #s145_FixClamp_T1;
   IF #s145_FixClamp THEN #StateNo := 145; END_IF;
END_REGION

REGION Network 28: Actions for STATE Num:145 Fix Clamp
   RUNG wire#powerrail
      Contact( #s145_FixClamp )
      Coil( #qFixClamp )
   END_RUNG
   // the same network as SCL:
   #qFixClamp := #s145_FixClamp;
END_REGION

REGION Network 29: Transition for STATE Num:146 Robot-2 All Alloys Pick Or Drop Operation over
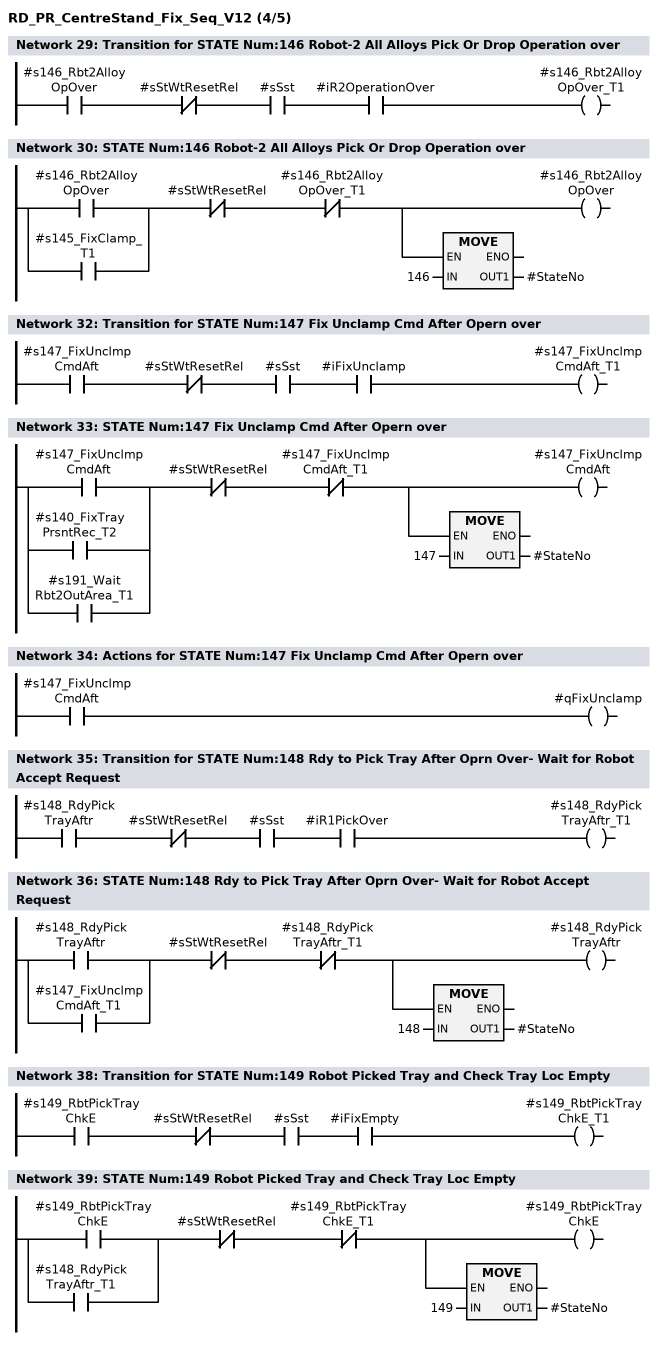
   RUNG wire#powerrail
      Contact( #s146_Rbt2AlloyOpOver )
      I_Contact( #sStWtResetRel )
      Contact( #sSst )
      Contact( #iR2OperationOver )
      Coil( #s146_Rbt2AlloyOpOver_T1 )
   END_RUNG
   // the same network as SCL:
   #s146_Rbt2AlloyOpOver_T1 := #s146_Rbt2AlloyOpOver AND NOT #sStWtResetRel AND #sSst AND #iR2OperationOver;
END_REGION

REGION Network 30: STATE Num:146 Robot-2 All Alloys Pick Or Drop Operation over
   RUNG wire#powerrail
      Contact( #s146_Rbt2AlloyOpOver )
      wire#w1
      I_Contact( #sStWtResetRel )
      I_Contact( #s146_Rbt2AlloyOpOver_T1 )
      wire#w2
      Coil( #s146_Rbt2AlloyOpOver )
   END_RUNG
   RUNG wire#powerrail
      Contact( #s145_FixClamp_T1 )
   END_RUNG wire#w1
   RUNG wire#w2
      { S7_GenerateENO := "TRUE" } Move(in := 146, out1 => #StateNo)
   END_RUNG
   // the same network as SCL:
   #s146_Rbt2AlloyOpOver := (#s146_Rbt2AlloyOpOver OR #s145_FixClamp_T1) AND NOT #sStWtResetRel AND NOT #s146_Rbt2AlloyOpOver_T1;
   IF #s146_Rbt2AlloyOpOver THEN #StateNo := 146; END_IF;
END_REGION

NETWORK
TITLE = Actions for STATE Num:146 Robot-2 All Alloys Pick Or Drop Operation over
      A     #s146_Rbt2AlloyOpOver;
      =     #qR2OperationStart;
      A     #s146_Rbt2AlloyOpOver;
      A     #iR2ServiceActivated;
      S     #iqR2ServiceActive;
      A     #s146_Rbt2AlloyOpOver;
      A     #iR2OperationOver;
      A     #iqR2ServiceActive;
      R     #iqR2ServiceActive;

REGION Network 32: Transition for STATE Num:147 Fix Unclamp Cmd After Opern over
   RUNG wire#powerrail
      Contact( #s147_FixUnclmpCmdAft )
      I_Contact( #sStWtResetRel )
      Contact( #sSst )
      Contact( #iFixUnclamp )
      Coil( #s147_FixUnclmpCmdAft_T1 )
   END_RUNG
   // the same network as SCL:
   #s147_FixUnclmpCmdAft_T1 := #s147_FixUnclmpCmdAft AND NOT #sStWtResetRel AND #sSst AND #iFixUnclamp;
END_REGION

REGION Network 33: STATE Num:147 Fix Unclamp Cmd After Opern over
   RUNG wire#powerrail
      Contact( #s147_FixUnclmpCmdAft )
      wire#w1
      I_Contact( #sStWtResetRel )
      I_Contact( #s147_FixUnclmpCmdAft_T1 )
      wire#w2
      Coil( #s147_FixUnclmpCmdAft )
   END_RUNG
   RUNG wire#powerrail
      Contact( #s140_FixTrayPrsntRec_T2 )
   END_RUNG wire#w1
   RUNG wire#powerrail
      Contact( #s191_WaitRbt2OutArea_T1 )
   END_RUNG wire#w1
   RUNG wire#w2
      { S7_GenerateENO := "TRUE" } Move(in := 147, out1 => #StateNo)
   END_RUNG
   // the same network as SCL:
   #s147_FixUnclmpCmdAft := (#s147_FixUnclmpCmdAft OR #s140_FixTrayPrsntRec_T2 OR #s191_WaitRbt2OutArea_T1) AND NOT #sStWtResetRel AND NOT #s147_FixUnclmpCmdAft_T1;
   IF #s147_FixUnclmpCmdAft THEN #StateNo := 147; END_IF;
END_REGION

REGION Network 34: Actions for STATE Num:147 Fix Unclamp Cmd After Opern over
   RUNG wire#powerrail
      Contact( #s147_FixUnclmpCmdAft )
      Coil( #qFixUnclamp )
   END_RUNG
   // the same network as SCL:
   #qFixUnclamp := #s147_FixUnclmpCmdAft;
END_REGION

REGION Network 35: Transition for STATE Num:148 Rdy to Pick Tray After Oprn Over- Wait for Robot Accept Request
   RUNG wire#powerrail
      Contact( #s148_RdyPickTrayAftr )
      I_Contact( #sStWtResetRel )
      Contact( #sSst )
      Contact( #iR1PickOver )
      Coil( #s148_RdyPickTrayAftr_T1 )
   END_RUNG
   // the same network as SCL:
   #s148_RdyPickTrayAftr_T1 := #s148_RdyPickTrayAftr AND NOT #sStWtResetRel AND #sSst AND #iR1PickOver;
END_REGION

REGION Network 36: STATE Num:148 Rdy to Pick Tray After Oprn Over- Wait for Robot Accept Request
   RUNG wire#powerrail
      Contact( #s148_RdyPickTrayAftr )
      wire#w1
      I_Contact( #sStWtResetRel )
      I_Contact( #s148_RdyPickTrayAftr_T1 )
      wire#w2
      Coil( #s148_RdyPickTrayAftr )
   END_RUNG
   RUNG wire#powerrail
      Contact( #s147_FixUnclmpCmdAft_T1 )
   END_RUNG wire#w1
   RUNG wire#w2
      { S7_GenerateENO := "TRUE" } Move(in := 148, out1 => #StateNo)
   END_RUNG
   // the same network as SCL:
   #s148_RdyPickTrayAftr := (#s148_RdyPickTrayAftr OR #s147_FixUnclmpCmdAft_T1) AND NOT #sStWtResetRel AND NOT #s148_RdyPickTrayAftr_T1;
   IF #s148_RdyPickTrayAftr THEN #StateNo := 148; END_IF;
END_REGION

NETWORK
TITLE = Actions for STATE Num:148 Rdy to Pick Tray After Oprn Over- Wait for Robot Accept Request
      A     #s148_RdyPickTrayAftr;
      =     #qR1ReadytoPickTray;
      A     #s148_RdyPickTrayAftr;
      A     #iR1PickOver;
      R     #iqR2ServiceCompleted;

REGION Network 38: Transition for STATE Num:149 Robot Picked Tray and Check Tray Loc Empty
   RUNG wire#powerrail
      Contact( #s149_RbtPickTrayChkE )
      I_Contact( #sStWtResetRel )
      Contact( #sSst )
      Contact( #iFixEmpty )
      Coil( #s149_RbtPickTrayChkE_T1 )
   END_RUNG
   // the same network as SCL:
   #s149_RbtPickTrayChkE_T1 := #s149_RbtPickTrayChkE AND NOT #sStWtResetRel AND #sSst AND #iFixEmpty;
END_REGION

REGION Network 39: STATE Num:149 Robot Picked Tray and Check Tray Loc Empty
   RUNG wire#powerrail
      Contact( #s149_RbtPickTrayChkE )
      wire#w1
      I_Contact( #sStWtResetRel )
      I_Contact( #s149_RbtPickTrayChkE_T1 )
      wire#w2
      Coil( #s149_RbtPickTrayChkE )
   END_RUNG
   RUNG wire#powerrail
      Contact( #s148_RdyPickTrayAftr_T1 )
   END_RUNG wire#w1
   RUNG wire#w2
      { S7_GenerateENO := "TRUE" } Move(in := 149, out1 => #StateNo)
   END_RUNG
   // the same network as SCL:
   #s149_RbtPickTrayChkE := (#s149_RbtPickTrayChkE OR #s148_RdyPickTrayAftr_T1) AND NOT #sStWtResetRel AND NOT #s149_RbtPickTrayChkE_T1;
   IF #s149_RbtPickTrayChkE THEN #StateNo := 149; END_IF;
END_REGION

REGION Network 40: Actions for STATE Num:149 Robot Picked Tray and Check Tray Loc Empty
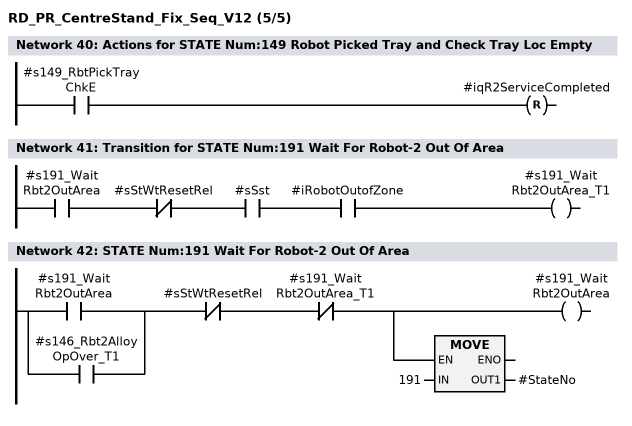
   RUNG wire#powerrail
      Contact( #s149_RbtPickTrayChkE )
      R_Coil( #iqR2ServiceCompleted )
   END_RUNG
   // the same network as SCL:
   IF #s149_RbtPickTrayChkE THEN #iqR2ServiceCompleted := FALSE; END_IF;
END_REGION

REGION Network 41: Transition for STATE Num:191 Wait For Robot-2 Out Of Area
   RUNG wire#powerrail
      Contact( #s191_WaitRbt2OutArea )
      I_Contact( #sStWtResetRel )
      Contact( #sSst )
      Contact( #iRobotOutofZone )
      Coil( #s191_WaitRbt2OutArea_T1 )
   END_RUNG
   // the same network as SCL:
   #s191_WaitRbt2OutArea_T1 := #s191_WaitRbt2OutArea AND NOT #sStWtResetRel AND #sSst AND #iRobotOutofZone;
END_REGION

REGION Network 42: STATE Num:191 Wait For Robot-2 Out Of Area
   RUNG wire#powerrail
      Contact( #s191_WaitRbt2OutArea )
      wire#w1
      I_Contact( #sStWtResetRel )
      I_Contact( #s191_WaitRbt2OutArea_T1 )
      wire#w2
      Coil( #s191_WaitRbt2OutArea )
   END_RUNG
   RUNG wire#powerrail
      Contact( #s146_Rbt2AlloyOpOver_T1 )
   END_RUNG wire#w1
   RUNG wire#w2
      { S7_GenerateENO := "TRUE" } Move(in := 191, out1 => #StateNo)
   END_RUNG
   // the same network as SCL:
   #s191_WaitRbt2OutArea := (#s191_WaitRbt2OutArea OR #s146_Rbt2AlloyOpOver_T1) AND NOT #sStWtResetRel AND NOT #s191_WaitRbt2OutArea_T1;
   IF #s191_WaitRbt2OutArea THEN #StateNo := 191; END_IF;
END_REGION
END_FUNCTION_BLOCK

